// TIA Portal project "PROYECTO PICK AND PLACE FUNCIONA" (V17)

(* hardware
DEVICE "S7-1200 station_1"  S7-1200 Station
   slot 0: "Rack_0"  S7-1200 Rack  Rack  V1.0
   slot 1: "PLC_1"  CPU 1214C AC/DC/Rly  6ES7 214-1BG40-0XB0  V4.5
DEVICE "Estación PC"  SIMATIC PC station
   slot 0: "Estación PC"  Rail  SIMATIC PC-Station  V1.0
      slot 125: "Stationmanager"  Station_Manager  V6.0.4
   slot 1: "IE general_1"  IE General  IE_CP  V8.2.0
      slot 1: "PROFINET interface"  IEGeneral.Interface.8.2.0
   slot 2: "HMI_RT_2"  WinCC RT Advanced  6AV2 104-0xxxx-xxxx  17.0.0.0
      slot 33792: "Interfaz del equipo"  Host interface
*)

// ===== PLC "PLC_1"  CPU 1214C AC/DC/Rly =====

VAR_GLOBAL   // PLC tag table "Tabla de variables estándar"
   "System_Byte" AT %MB1 : Byte;
   "FirstScan" AT %M1.0 : Bool;
   "DiagStatusUpdate" AT %M1.1 : Bool;
   "AlwaysTRUE" AT %M1.2 : Bool;
   "AlwaysFALSE" AT %M1.3 : Bool;
   "Tag_1" AT %M700.3 : Bool;
   "Tag_2" AT %M700.4 : Bool;
   "Tag_3" AT %M900.0 : Bool;
   "Tag_4" AT %M900.1 : Bool;
   "Tag_5" AT %M900.5 : Bool;
   "MARCA_VENTOSA_V3" AT %M3000.0 : Bool;
   "Tag_6" AT %M8765.0 : Bool;
   "MARCA VACIA" AT %M3214.0 : Bool;
   "MARCA_VACIAA" AT %M4500.0 : Bool;
   "Tag_7" AT %MW5000 : Word;
   "Tag_8" AT %MD5000 : DWord;
   "RESET_CTU" AT %M5000.0 : Bool;
   "Tag_9" AT %MD5010 : DInt;
   "Tag_10" AT %M763.3 : Bool;
   "Tag_11" AT %M668.2 : Bool;
   "Tag_12" AT %M668.3 : Bool;
   "Tag_13" AT %M996.0 : Bool;
   "Tag_14" AT %M1200.0 : Bool;
   "Tag_15" AT %M1200.2 : Bool;
   "POSICIÓN 1" AT %M543.0 : Bool;
   "POSICIÓN 2" AT %M543.1 : Bool;
   "POSICIÓN 3" AT %M543.2 : Bool;
   "POSICIÓN 4" AT %M543.3 : Bool;
   "POSICIÓN 5" AT %M543.4 : Bool;
   "POSICIÓN 6" AT %M543.5 : Bool;
   "POSICIÓN 7" AT %M543.6 : Bool;
   "POSICIÓN 8" AT %M543.7 : Bool;
   "POSICIÓN 9" AT %M544.0 : Bool;
   "POSICIÓN 10" AT %M544.1 : Bool;
   "Tag_16" AT %M545.3 : Bool;
   "VALOR_PROCESO_ENTRADA" AT %QW15 : Int;
   "VALOR_PROCESO_SALIDA" AT %QW20 : Int;
END_VAR

VAR_GLOBAL   // PLC tag table "ENTRADAS Y SALIDAS"
   "PULSADOR_S1" AT %I0.0 : Bool;
   "PULSADOR_S2" AT %I0.1 : Bool;
   "SELECTOR_S3" AT %I0.2 : Bool;
   "PULSADOR_S4" AT %I0.3 : Bool;
   "DETECTOR_B1" AT %I0.4 : Bool;
   "DETECTOR_B2" AT %I0.5 : Bool;
   "DETECTOR_B3" AT %I0.6 : Bool;
   "DETECTOR_B4" AT %I0.7 : Bool;
   "DETECTOR_B5" AT %I1.0 : Bool;
   "E.VALVULA_MB1(B+)" AT %Q0.0 : Bool;
   "E.VALVULA_MB2(A+)" AT %Q0.1 : Bool;
   "CINTA1_KM1" AT %Q0.2 : Bool;
   "CINTA2_KM2" AT %Q0.3 : Bool;
   "VENTOSA_V1" AT %Q0.4 : Bool;
   "PILOTO_H2" AT %Q0.5 : Bool;
   "PILOTO_H1" AT %Q0.6 : Bool;
   "PILOTO_H3(AUTO)" AT %Q0.7 : Bool;
   "SELECTOR_S7" AT %I1.2 : Bool;
   "CINTA3_KM3" AT %Q1.0 : Bool;
   "CINTA4_KM4" AT %Q1.1 : Bool;
   "CINTA5_KM5" AT %Q1.2 : Bool;
   "CINTA6_KM6" AT %Q1.3 : Bool;
   "BARRERA1_KM7" AT %Q1.4 : Bool;
   "DETECTOR_B8=B3" AT %I1.4 : Bool;
   "DETECTOR C+_B9=B7" AT %I1.5 : Bool;
   "DETECTOR D+_B10=B6" AT %I1.6 : Bool;
   "DETECTOR_B11=B1" AT %I1.7 : Bool;
   "DETECTOR_B12=B4" AT %I2.0 : Bool;
   "DETECTOR_B13=B2" AT %I2.1 : Bool;
   "DETECTOR_B14=B5" AT %I2.2 : Bool;
   "BARRERA2_KM8" AT %Q1.5 : Bool;
   "PILOTO_H6(ROJO)" AT %Q2.0 : Bool;
   "PILOTO_H4(VERDE)" AT %Q2.1 : Bool;
   "PILOTO_H5(AMARILLO)" AT %Q2.2 : Bool;
   "M.MANUA2_S9" AT %I2.3 : Bool;
   "AUTO2_S10" AT %I2.4 : Bool;
   "MARCHA2_S5" AT %I2.5 : Bool;
   "PULSADOR_MANUAL_S6" AT %I2.6 : Bool;
   "PARO2_S8" AT %I2.7 : Bool;
   "PILOTO_H12=H1" AT %Q2.3 : Bool;
   "PILOTO_H7=H2" AT %Q2.4 : Bool;
   "PILOTO_H8=H3" AT %Q2.5 : Bool;
   "CINTA7_KM9=KM3" AT %Q2.6 : Bool;
   "PILOTO_H9=H4" AT %Q2.7 : Bool;
   "PILOTO_H10=H5" AT %Q3.0 : Bool;
   "PILOTO_H11=H6" AT %Q3.1 : Bool;
   "CILINDRO_C=A" AT %Q1.6 : Bool;
   "CILINDRO_D=B" AT %Q1.7 : Bool;
   "VENTOSA_V2" AT %Q3.2 : Bool;
   "FC1_E+" AT %I3.0 : Bool;
   "CILINDRO E" AT %Q5.0 : Bool;
   "FC2_E-" AT %I3.1 : Bool;
   "CÁMARA1_B15(AZUL)" AT %I3.2 : Bool;
   "CÁMARA2_B16(VERDE)" AT %I3.3 : Bool;
   "FC4_F+" AT %I3.4 : Bool;
   "FC5_G-" AT %I3.5 : Bool;
   "FC6_G+" AT %I3.6 : Bool;
   "FC3_F-" AT %I3.7 : Bool;
   "CILINDRO F" AT %Q5.1 : Bool;
   "CILINDRO G" AT %QD38 : DWord;
   "CINTA8_KM10" AT %Q3.3 : Bool;
   "PILOTOEMERGENCIA_H13" AT %Q3.4 : Bool;
   "SETAEMERGENCIA_S12" AT %I4.0 : Bool;
   "RESET1_S11" AT %I4.1 : Bool;
   "RESET2_S14" AT %I4.2 : Bool;
   "SETAEMERGENCIA2_S13" AT %I4.3 : Bool;
   "PILOTOEMERGENCIA2_H14" AT %Q3.5 : Bool;
   "DETECTOR_B15" AT %I4.4 : Bool;
   "ROBOT_OCUPADO_B16" AT %I4.5 : Bool;
   "ROBOT_ERROR_B17" AT %I4.6 : Bool;
   "ACTIVACIÓN_ROBOT" AT %Q3.6 : Bool;
   "DETECTOR_B21(INICIO P.AZUL)" AT %I4.7 : Bool;
   "DETECTOR_B22(FINAL P.AZUL)" AT %I5.0 : Bool;
   "CINTA9_KM11(BASE AZUL)" AT %Q3.7 : Bool;
   "CINTA10_KM12(BASE AZUL)" AT %Q4.0 : Bool;
   "CINTA11_KM13(BASE AZUL)" AT %Q4.1 : Bool;
   "BARRERA3_KM14(BASE AZUL)" AT %Q4.2 : Bool;
   "EJE_X1" AT %QD42 : Real;
   "EJE_Y1" AT %QD46 : Real;
   "EJE_Z1" AT %QD50 : Real;
   "VENTOSA_V3" AT %Q4.3 : Bool;
   "CINTA12_KM15(BASE VERDE)" AT %Q4.4 : Bool;
   "CINTA13_KM16(BASE VERDE)" AT %Q4.5 : Bool;
   "CINTA14_KM17(BASE VERDE)" AT %Q4.6 : Bool;
   "BARRERA4_KM18" AT %Q4.7 : Bool;
   "DETECTOR_B23(INICIO BASE VERDE)" AT %I5.1 : Bool;
   "DETECTOR_B24(FINAL BASE VERDE)" AT %I5.2 : Bool;
   "EJE_X2" AT %QD34 : Real;
   "EJE_Y2" AT %QD54 : Real;
   "EJE_Z2" AT %QD58 : Real;
   "VENTOSA_V4" AT %Q5.2 : Bool;
   "CINTA15_KM19" AT %Q5.3 : Bool;
   "CINTA16_KM20" AT %Q5.4 : Bool;
   "CINTA17_KM21" AT %Q5.5 : Bool;
   "CINTA18_KM22" AT %Q5.6 : Bool;
   "CINTA19_KM23" AT %Q5.7 : Bool;
   "CINTA20_KM24" AT %Q6.0 : Bool;
   "UÑASATRAS_KM25" AT %Q6.1 : Bool;
   "VAGÓN_ARRIBA_KM26" AT %Q6.2 : Bool;
   "SELECCION POSICIÓN" AT %QD30 : DInt;
   "DETECTOR_B25" AT %I5.3 : Bool;
   "DETECTOR_B26" AT %I5.4 : Bool;
   "SALIDA BASES" AT %Q6.3 : Bool;
   "SALIDA PALET_AZUL" AT %Q6.4 : Bool;
   "UÑAS_ALANTE_KM27" AT %Q6.5 : Bool;
   "CINTA21_KM28" AT %Q6.6 : Bool;
   "CINTA22_KM29" AT %Q6.7 : Bool;
   "CINTA23_KM30" AT %Q7.0 : Bool;
   "CINTA24_KM31" AT %Q7.1 : Bool;
   "CINTA25_KM32" AT %Q7.2 : Bool;
   "CINTA26_KM33" AT %Q7.3 : Bool;
   "DETECTOR_B27" AT %I5.5 : Bool;
   "DETECTOR_B28" AT %I5.6 : Bool;
   "SALIDA_PALET_VERDE" AT %Q7.4 : Bool;
   "VALOR_CONTADOR" AT %IW6 : Int;
   "MARCAA_VACIIA" AT %M730.0 : Bool;
END_VAR

VAR_GLOBAL   // PLC tag table "ETAPAS"
   "ETAPA_1" AT %M10.1 : Bool;
   "ETAPA_2" AT %M10.2 : Bool;
   "ETAPA_3" AT %M10.3 : Bool;
   "ETAPA_4" AT %M10.4 : Bool;
   "ETAPA_5" AT %M10.5 : Bool;
   "ETAPA_6" AT %M10.6 : Bool;
   "ETAPA_7" AT %M10.7 : Bool;
   "ETAPA_12" AT %M11.0 : Bool;
   "ETAPA_13" AT %M11.1 : Bool;
   "ETAPA_14" AT %M11.2 : Bool;
   "ETAPA_15" AT %M11.3 : Bool;
   "ETAPA_16" AT %M11.4 : Bool;
   "ETAPA_17" AT %M11.5 : Bool;
   "ETAPA_0" AT %M10.0 : Bool;
   "ETAPA_100" AT %M11.6 : Bool;
   "ETAPA_101" AT %M11.7 : Bool;
   "ETAPA_50" AT %M12.0 : Bool;
   "ETAPA_51" AT %M12.1 : Bool;
   "ETAPA_54" AT %M12.2 : Bool;
   "ETAPA_55" AT %M12.3 : Bool;
   "ETAPA_56" AT %M12.4 : Bool;
   "ETAPA_57" AT %M12.5 : Bool;
   "ETAPA_58" AT %M12.6 : Bool;
   "ETAPA_59" AT %M12.7 : Bool;
   "ETAPA_62" AT %M13.0 : Bool;
   "ETAPA_63" AT %M13.1 : Bool;
   "ETAPA_64" AT %M13.2 : Bool;
   "ETAPA_65" AT %M13.3 : Bool;
   "ETAPA_66" AT %M13.4 : Bool;
   "ETAPA_67" AT %M13.5 : Bool;
   "ETAPA_52" AT %M14.0 : Bool;
   "ETAPA_53" AT %M14.1 : Bool;
   "ETAPA_60" AT %M14.2 : Bool;
   "ETAPA_61" AT %M14.3 : Bool;
   "ETAPA_8" AT %M14.4 : Bool;
   "ETAPA_9" AT %M14.5 : Bool;
   "ETAPA_18" AT %M14.6 : Bool;
   "ETAPA_19" AT %M14.7 : Bool;
   "ETAPA_20" AT %M15.1 : Bool;
   "ETAPA_21" AT %M15.2 : Bool;
   "ETAPA _10" AT %M15.3 : Bool;
   "ETAPA_11" AT %M15.4 : Bool;
   "ETAPA_120" AT %M15.5 : Bool;
   "ETAPA_121" AT %M23.0 : Bool;
   "ETAPA_140" AT %M15.7 : Bool;
   "ETAPA_141" AT %M16.0 : Bool;
   "ETAPA_160" AT %M16.1 : Bool;
   "ETAPA_161" AT %M16.2 : Bool;
   "ETAPA_200" AT %M16.3 : Bool;
   "ETAPA_201" AT %M16.4 : Bool;
   "ETAPA_202" AT %M16.5 : Bool;
   "ETAPA_203" AT %M16.6 : Bool;
   "ETAPA_204" AT %M16.7 : Bool;
   "ETAPA_205" AT %M17.0 : Bool;
   "ETAPA_206" AT %M17.1 : Bool;
   "ETAPA_207" AT %M17.2 : Bool;
   "ETAPA_208" AT %M17.3 : Bool;
   "ETAPA_209" AT %M17.4 : Bool;
   "ETAPA_210" AT %M17.5 : Bool;
   "ETAPA_211" AT %M17.6 : Bool;
   "ETAPA_212" AT %M17.7 : Bool;
   "ETAPA_213" AT %M18.0 : Bool;
   "ETAPA_214" AT %M18.1 : Bool;
   "ETAPA_215" AT %M18.2 : Bool;
   "ETAPA_216" AT %M18.3 : Bool;
   "ETAPA_217" AT %M18.4 : Bool;
   "ETAPA_218" AT %M18.5 : Bool;
   "ETAPA_250" AT %M18.6 : Bool;
   "ETAPA_251" AT %M18.7 : Bool;
   "ETAPA_252" AT %M19.0 : Bool;
   "ETAPA_253" AT %M19.1 : Bool;
   "ETAPA_254" AT %M19.2 : Bool;
   "ETAPA_255" AT %M19.3 : Bool;
   "ETAPA_256" AT %M19.4 : Bool;
   "ETAPA_257" AT %M19.5 : Bool;
   "ETAPA_258" AT %M19.6 : Bool;
   "ETAPA_259" AT %M19.7 : Bool;
   "ETAPA_260" AT %M20.0 : Bool;
   "ETAPA_261" AT %M20.1 : Bool;
   "ETAPA_262" AT %M20.2 : Bool;
   "ETAPA_263" AT %M20.3 : Bool;
   "ETAPA_264" AT %M20.4 : Bool;
   "ETAPA_265" AT %M20.5 : Bool;
   "ETAPA_266" AT %M20.6 : Bool;
END_VAR

// folder: System blocks/Program resources

DATA_BLOCK "TEMPORIZADOR 1"   // DB1
{ S7_Optimized_Access := 'TRUE' }
AUTHOR : Simatic
FAMILY : IEC
NAME : IEC_TMR
VERSION : 1.0
// stored: InstanceOfName IEC_TIMER
"IEC_TIMER"
BEGIN
END_DATA_BLOCK

DATA_BLOCK "TEMPORIZADOR 2"   // DB2
{ S7_Optimized_Access := 'TRUE' }
AUTHOR : Simatic
FAMILY : IEC
NAME : IEC_TMR
VERSION : 1.0
// stored: InstanceOfName IEC_TIMER
"IEC_TIMER"
BEGIN
END_DATA_BLOCK

DATA_BLOCK "TEMPORIZADOR 3"   // DB3
{ S7_Optimized_Access := 'TRUE' }
AUTHOR : Simatic
FAMILY : IEC
NAME : IEC_TMR
VERSION : 1.0
// stored: InstanceOfName IEC_TIMER
"IEC_TIMER"
BEGIN
END_DATA_BLOCK

DATA_BLOCK "TEMPORIZADOR 4"   // DB4
{ S7_Optimized_Access := 'TRUE' }
AUTHOR : Simatic
FAMILY : IEC
NAME : IEC_TMR
VERSION : 1.0
// stored: InstanceOfName IEC_TIMER
"IEC_TIMER"
BEGIN
END_DATA_BLOCK

DATA_BLOCK "TEMPORIZADOR 5"   // DB5
{ S7_Optimized_Access := 'TRUE' }
AUTHOR : Simatic
FAMILY : IEC
NAME : IEC_TMR
VERSION : 1.0
// stored: InstanceOfName IEC_TIMER
"IEC_TIMER"
BEGIN
END_DATA_BLOCK

DATA_BLOCK "TEMPORIZADOR 6"   // DB6
{ S7_Optimized_Access := 'TRUE' }
AUTHOR : Simatic
FAMILY : IEC
NAME : IEC_TMR
VERSION : 1.0
// stored: InstanceOfName IEC_TIMER
"IEC_TIMER"
BEGIN
END_DATA_BLOCK

DATA_BLOCK "TEMPORIZADOR 10"   // DB7
{ S7_Optimized_Access := 'TRUE' }
AUTHOR : Simatic
FAMILY : IEC
NAME : IEC_TMR
VERSION : 1.0
// stored: InstanceOfName IEC_TIMER
"IEC_TIMER"
BEGIN
END_DATA_BLOCK

DATA_BLOCK "TEMPORIZADOR 8"   // DB8
{ S7_Optimized_Access := 'TRUE' }
AUTHOR : Simatic
FAMILY : IEC
NAME : IEC_TMR
VERSION : 1.0
// stored: InstanceOfName IEC_TIMER
"IEC_TIMER"
BEGIN
END_DATA_BLOCK

DATA_BLOCK "TEMPORIZADOR 13"   // DB9
{ S7_Optimized_Access := 'TRUE' }
AUTHOR : Simatic
FAMILY : IEC
NAME : IEC_TMR
VERSION : 1.0
// stored: InstanceOfName IEC_TIMER
"IEC_TIMER"
BEGIN
END_DATA_BLOCK

DATA_BLOCK "TEMPORIZADOR 15"   // DB10
{ S7_Optimized_Access := 'TRUE' }
AUTHOR : Simatic
FAMILY : IEC
NAME : IEC_TMR
VERSION : 1.0
// stored: InstanceOfName IEC_TIMER
"IEC_TIMER"
BEGIN
END_DATA_BLOCK

DATA_BLOCK "TEMPORIZADOR 11"   // DB11
{ S7_Optimized_Access := 'TRUE' }
AUTHOR : Simatic
FAMILY : IEC
NAME : IEC_TMR
VERSION : 1.0
// stored: InstanceOfName IEC_TIMER
"IEC_TIMER"
BEGIN
END_DATA_BLOCK

DATA_BLOCK "TEMPORIZADOR 14"   // DB12
{ S7_Optimized_Access := 'TRUE' }
AUTHOR : Simatic
FAMILY : IEC
NAME : IEC_TMR
VERSION : 1.0
// stored: InstanceOfName IEC_TIMER
"IEC_TIMER"
BEGIN
END_DATA_BLOCK

DATA_BLOCK "TEMPORIZADOR 7"   // DB13
{ S7_Optimized_Access := 'TRUE' }
AUTHOR : Simatic
FAMILY : IEC
NAME : IEC_TMR
VERSION : 1.0
// stored: InstanceOfName IEC_TIMER
"IEC_TIMER"
BEGIN
END_DATA_BLOCK

DATA_BLOCK "TEMPORIZADOR 16"   // DB14
{ S7_Optimized_Access := 'TRUE' }
AUTHOR : Simatic
FAMILY : IEC
NAME : IEC_TMR
VERSION : 1.0
// stored: InstanceOfName IEC_TIMER
"IEC_TIMER"
BEGIN
END_DATA_BLOCK

DATA_BLOCK "TEMPORIZADOR 17"   // DB15
{ S7_Optimized_Access := 'TRUE' }
AUTHOR : Simatic
FAMILY : IEC
NAME : IEC_TMR
VERSION : 1.0
// stored: InstanceOfName IEC_TIMER
"IEC_TIMER"
BEGIN
END_DATA_BLOCK

DATA_BLOCK "TEMPORIZADOR 18"   // DB16
{ S7_Optimized_Access := 'TRUE' }
AUTHOR : Simatic
FAMILY : IEC
NAME : IEC_TMR
VERSION : 1.0
// stored: InstanceOfName IEC_TIMER
"IEC_TIMER"
BEGIN
END_DATA_BLOCK

DATA_BLOCK "TEMPORIZADOR 19"   // DB17
{ S7_Optimized_Access := 'TRUE' }
AUTHOR : Simatic
FAMILY : IEC
NAME : IEC_TMR
VERSION : 1.0
// stored: InstanceOfName IEC_TIMER
"IEC_TIMER"
BEGIN
END_DATA_BLOCK

DATA_BLOCK "TEMPORIZADOR 20"   // DB18
{ S7_Optimized_Access := 'TRUE' }
AUTHOR : Simatic
FAMILY : IEC
NAME : IEC_TMR
VERSION : 1.0
// stored: InstanceOfName IEC_TIMER
"IEC_TIMER"
BEGIN
END_DATA_BLOCK

DATA_BLOCK "TEMPORIZADOR 21"   // DB19
{ S7_Optimized_Access := 'TRUE' }
AUTHOR : Simatic
FAMILY : IEC
NAME : IEC_TMR
VERSION : 1.0
// stored: InstanceOfName IEC_TIMER
"IEC_TIMER"
BEGIN
END_DATA_BLOCK

DATA_BLOCK "TEMPORIZADOR 22"   // DB20
{ S7_Optimized_Access := 'TRUE' }
AUTHOR : Simatic
FAMILY : IEC
NAME : IEC_TMR
VERSION : 1.0
// stored: InstanceOfName IEC_TIMER
"IEC_TIMER"
BEGIN
END_DATA_BLOCK

DATA_BLOCK "IEC_Timer_0_DB"   // DB21
{ S7_Optimized_Access := 'TRUE' }
AUTHOR : Simatic
FAMILY : IEC
NAME : IEC_TMR
VERSION : 1.0
// stored: InstanceOfName IEC_TIMER
"IEC_TIMER"
BEGIN
END_DATA_BLOCK

DATA_BLOCK "TEMPORIZADOR 23"   // DB22
{ S7_Optimized_Access := 'TRUE' }
AUTHOR : Simatic
FAMILY : IEC
NAME : IEC_TMR
VERSION : 1.0
// stored: InstanceOfName IEC_TIMER
"IEC_TIMER"
BEGIN
END_DATA_BLOCK

DATA_BLOCK "TEMPORIZADOR 24"   // DB23
{ S7_Optimized_Access := 'TRUE' }
AUTHOR : Simatic
FAMILY : IEC
NAME : IEC_TMR
VERSION : 1.0
// stored: InstanceOfName IEC_TIMER
"IEC_TIMER"
BEGIN
END_DATA_BLOCK

DATA_BLOCK "TEMPORIZADOR 25"   // DB24
{ S7_Optimized_Access := 'TRUE' }
AUTHOR : Simatic
FAMILY : IEC
NAME : IEC_TMR
VERSION : 1.0
// stored: InstanceOfName IEC_TIMER
"IEC_TIMER"
BEGIN
END_DATA_BLOCK

DATA_BLOCK "TEMPORIZADOR 26"   // DB25
{ S7_Optimized_Access := 'TRUE' }
AUTHOR : Simatic
FAMILY : IEC
NAME : IEC_TMR
VERSION : 1.0
// stored: InstanceOfName IEC_TIMER
"IEC_TIMER"
BEGIN
END_DATA_BLOCK

DATA_BLOCK "TEMPORIZADOR 27"   // DB26
{ S7_Optimized_Access := 'TRUE' }
AUTHOR : Simatic
FAMILY : IEC
NAME : IEC_TMR
VERSION : 1.0
// stored: InstanceOfName IEC_TIMER
"IEC_TIMER"
BEGIN
END_DATA_BLOCK

DATA_BLOCK "TEMPORIZADOR 28"   // DB27
{ S7_Optimized_Access := 'TRUE' }
AUTHOR : Simatic
FAMILY : IEC
NAME : IEC_TMR
VERSION : 1.0
// stored: InstanceOfName IEC_TIMER
"IEC_TIMER"
BEGIN
END_DATA_BLOCK

DATA_BLOCK "TEMPORIZADOR 29"   // DB28
{ S7_Optimized_Access := 'TRUE' }
AUTHOR : Simatic
FAMILY : IEC
NAME : IEC_TMR
VERSION : 1.0
// stored: InstanceOfName IEC_TIMER
"IEC_TIMER"
BEGIN
END_DATA_BLOCK

DATA_BLOCK "TEMPORIZADOR 30"   // DB29
{ S7_Optimized_Access := 'TRUE' }
AUTHOR : Simatic
FAMILY : IEC
NAME : IEC_TMR
VERSION : 1.0
// stored: InstanceOfName IEC_TIMER
"IEC_TIMER"
BEGIN
END_DATA_BLOCK

DATA_BLOCK "TEMPORIZADOR 31"   // DB30
{ S7_Optimized_Access := 'TRUE' }
AUTHOR : Simatic
FAMILY : IEC
NAME : IEC_TMR
VERSION : 1.0
// stored: InstanceOfName IEC_TIMER
"IEC_TIMER"
BEGIN
END_DATA_BLOCK

DATA_BLOCK "TEMPORIZADOR 32"   // DB31
{ S7_Optimized_Access := 'TRUE' }
AUTHOR : Simatic
FAMILY : IEC
NAME : IEC_TMR
VERSION : 1.0
// stored: InstanceOfName IEC_TIMER
"IEC_TIMER"
BEGIN
END_DATA_BLOCK

DATA_BLOCK "TEMPORIZADOR 33"   // DB32
{ S7_Optimized_Access := 'TRUE' }
AUTHOR : Simatic
FAMILY : IEC
NAME : IEC_TMR
VERSION : 1.0
// stored: InstanceOfName IEC_TIMER
"IEC_TIMER"
BEGIN
END_DATA_BLOCK

DATA_BLOCK "TEMPORIZADOR 34"   // DB33
{ S7_Optimized_Access := 'TRUE' }
AUTHOR : Simatic
FAMILY : IEC
NAME : IEC_TMR
VERSION : 1.0
// stored: InstanceOfName IEC_TIMER
"IEC_TIMER"
BEGIN
END_DATA_BLOCK

DATA_BLOCK "TEMPORIZADOR 35"   // DB34
{ S7_Optimized_Access := 'TRUE' }
AUTHOR : Simatic
FAMILY : IEC
NAME : IEC_TMR
VERSION : 1.0
// stored: InstanceOfName IEC_TIMER
"IEC_TIMER"
BEGIN
END_DATA_BLOCK

DATA_BLOCK "TEMPORIZADOR 36"   // DB35
{ S7_Optimized_Access := 'TRUE' }
AUTHOR : Simatic
FAMILY : IEC
NAME : IEC_TMR
VERSION : 1.0
// stored: InstanceOfName IEC_TIMER
"IEC_TIMER"
BEGIN
END_DATA_BLOCK

DATA_BLOCK "TEMPORIZADOR 37"   // DB36
{ S7_Optimized_Access := 'TRUE' }
AUTHOR : Simatic
FAMILY : IEC
NAME : IEC_TMR
VERSION : 1.0
// stored: InstanceOfName IEC_TIMER
"IEC_TIMER"
BEGIN
END_DATA_BLOCK

DATA_BLOCK "IEC_Timer_0_DB_1"   // DB37
{ S7_Optimized_Access := 'TRUE' }
AUTHOR : Simatic
FAMILY : IEC
NAME : IEC_TMR
VERSION : 1.0
// stored: InstanceOfName IEC_TIMER
"IEC_TIMER"
BEGIN
END_DATA_BLOCK

DATA_BLOCK "IEC_Counter_0_DB_1"   // DB38
{ S7_Optimized_Access := 'TRUE' }
AUTHOR : Simatic
FAMILY : IEC
NAME : CNTR
VERSION : 1.0
// stored: InstanceOfName IEC_COUNTER
"IEC_COUNTER"
BEGIN
END_DATA_BLOCK

DATA_BLOCK "IEC_Timer_0_DB_2"   // DB39
{ S7_Optimized_Access := 'TRUE' }
AUTHOR : Simatic
FAMILY : IEC
NAME : IEC_TMR
VERSION : 1.0
// stored: InstanceOfName IEC_TIMER
"IEC_TIMER"
BEGIN
END_DATA_BLOCK

DATA_BLOCK "IEC_Timer_0_DB_3"   // DB40
{ S7_Optimized_Access := 'TRUE' }
AUTHOR : Simatic
FAMILY : IEC
NAME : IEC_TMR
VERSION : 1.0
// stored: InstanceOfName IEC_TIMER
"IEC_TIMER"
BEGIN
END_DATA_BLOCK

DATA_BLOCK "TEMPORIZADOR 38"   // DB41
{ S7_Optimized_Access := 'TRUE' }
AUTHOR : Simatic
FAMILY : IEC
NAME : IEC_TMR
VERSION : 1.0
// stored: InstanceOfName IEC_TIMER
"IEC_TIMER"
BEGIN
END_DATA_BLOCK

DATA_BLOCK "TEMPORIZADOR 39"   // DB42
{ S7_Optimized_Access := 'TRUE' }
AUTHOR : Simatic
FAMILY : IEC
NAME : IEC_TMR
VERSION : 1.0
// stored: InstanceOfName IEC_TIMER
"IEC_TIMER"
BEGIN
END_DATA_BLOCK

DATA_BLOCK "IEC_Timer_0_DB_4"   // DB43
{ S7_Optimized_Access := 'TRUE' }
AUTHOR : Simatic
FAMILY : IEC
NAME : IEC_TMR
VERSION : 1.0
// stored: InstanceOfName IEC_TIMER
"IEC_TIMER"
BEGIN
END_DATA_BLOCK

DATA_BLOCK "IEC_Timer_0_DB_5"   // DB44
{ S7_Optimized_Access := 'TRUE' }
AUTHOR : Simatic
FAMILY : IEC
NAME : IEC_TMR
VERSION : 1.0
// stored: InstanceOfName IEC_TIMER
"IEC_TIMER"
BEGIN
END_DATA_BLOCK

DATA_BLOCK "TEMPORIZADOR 40"   // DB45
{ S7_Optimized_Access := 'TRUE' }
AUTHOR : Simatic
FAMILY : IEC
NAME : IEC_TMR
VERSION : 1.0
// stored: InstanceOfName IEC_TIMER
"IEC_TIMER"
BEGIN
END_DATA_BLOCK

DATA_BLOCK "TEMPORIZADOR 41"   // DB46
{ S7_Optimized_Access := 'TRUE' }
AUTHOR : Simatic
FAMILY : IEC
NAME : IEC_TMR
VERSION : 1.0
// stored: InstanceOfName IEC_TIMER
"IEC_TIMER"
BEGIN
END_DATA_BLOCK

DATA_BLOCK "TEMPORIZADOR 42"   // DB47
{ S7_Optimized_Access := 'TRUE' }
AUTHOR : Simatic
FAMILY : IEC
NAME : IEC_TMR
VERSION : 1.0
// stored: InstanceOfName IEC_TIMER
"IEC_TIMER"
BEGIN
END_DATA_BLOCK

DATA_BLOCK "TEMPORIZADOR 43"   // DB48
{ S7_Optimized_Access := 'TRUE' }
AUTHOR : Simatic
FAMILY : IEC
NAME : IEC_TMR
VERSION : 1.0
// stored: InstanceOfName IEC_TIMER
"IEC_TIMER"
BEGIN
END_DATA_BLOCK

DATA_BLOCK "TEMPORIZADOR 44"   // DB49
{ S7_Optimized_Access := 'TRUE' }
AUTHOR : Simatic
FAMILY : IEC
NAME : IEC_TMR
VERSION : 1.0
// stored: InstanceOfName IEC_TIMER
"IEC_TIMER"
BEGIN
END_DATA_BLOCK

DATA_BLOCK "TEMPORIZADOR 45"   // DB50
{ S7_Optimized_Access := 'TRUE' }
AUTHOR : Simatic
FAMILY : IEC
NAME : IEC_TMR
VERSION : 1.0
// stored: InstanceOfName IEC_TIMER
"IEC_TIMER"
BEGIN
END_DATA_BLOCK

// folder: (top level)

FUNCTION "FC_SECUENCIA SALIDA PARTE 1" : Void   // FC1, LAD
TITLE = PROGRAMACIÓN DEL PROCESO INDUSTRIAL
{ S7_Optimized_Access := 'TRUE' }
VERSION : 0.1
// ESTE BLOQUE MUESTRA LA PROGRAMACIÓN DE LA SECUENCIA DEL PROCESO INDUSTRIAL, DESDE QUE SALE DEL ROBOT HASTA QUE PASA LAS CÁMARAS DE VISIÓN DE COLORES
   VAR_TEMP   // added for the SCL form of the ladder/FBD networks
      _w1 : Bool;
      _w2 : Bool;
      _w3 : Bool;
      _w4 : Bool;
      _w5 : Bool;
   END_VAR
BEGIN

REGION Network 1: SET EN LA ETAPA 0
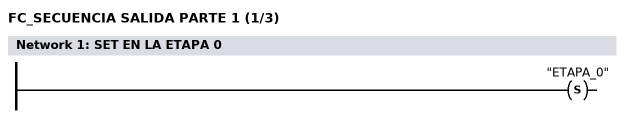
   RUNG wire#powerrail
      S_Coil( "ETAPA_0" )
   END_RUNG
   // the same network as SCL:
   "ETAPA_0" := TRUE;
END_REGION

REGION Network 2: PROGRAMACIÓN DE LA SECUENCIA EN MODO AUTOMÁTICO
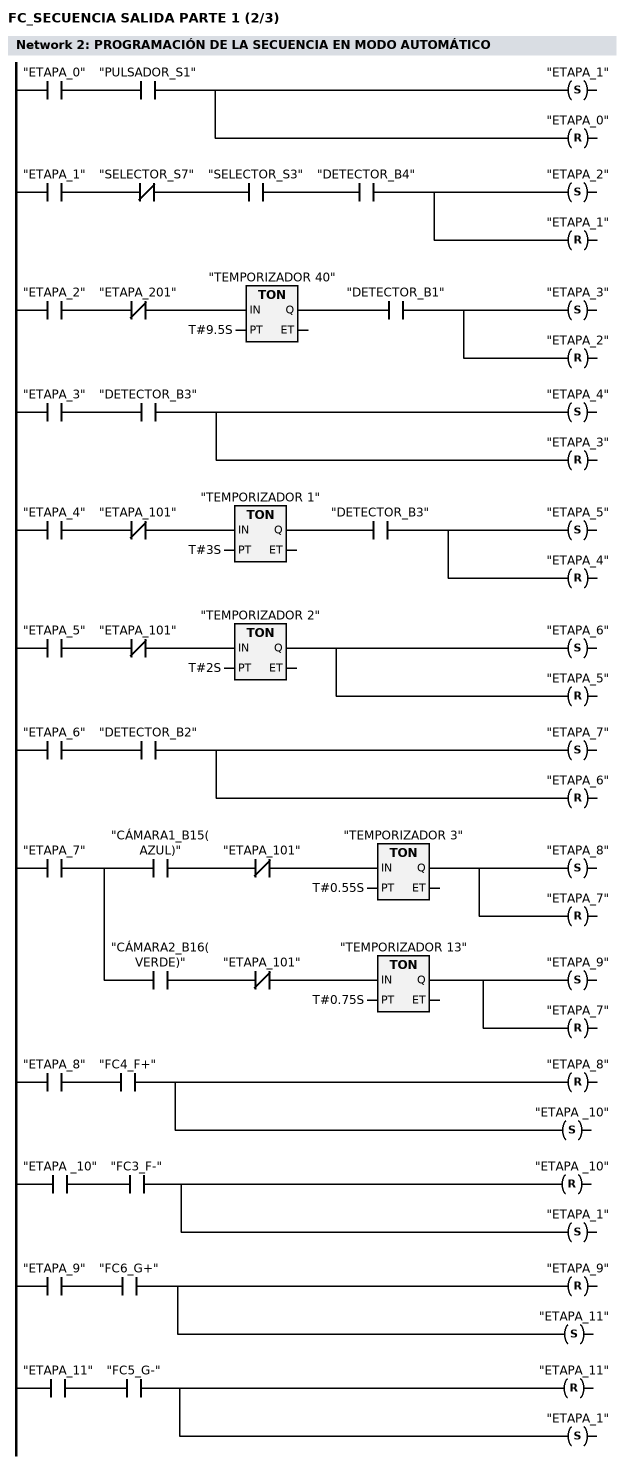
   IF "ETAPA_0" AND "PULSADOR_S1" THEN
       "ETAPA_1" := TRUE;
       "ETAPA_0" := FALSE;
   END_IF;
   IF "ETAPA_1" AND NOT "SELECTOR_S7" AND "SELECTOR_S3" AND "DETECTOR_B4" THEN
       "ETAPA_2" := TRUE;
       "ETAPA_1" := FALSE;
   END_IF;
   "TEMPORIZADOR 40".TON(IN := "ETAPA_2" AND NOT "ETAPA_201", PT := T#9.5S);
   IF "TEMPORIZADOR 40".Q AND "DETECTOR_B1" THEN
       "ETAPA_3" := TRUE;
       "ETAPA_2" := FALSE;
   END_IF;
   IF "ETAPA_3" AND "DETECTOR_B3" THEN
       "ETAPA_4" := TRUE;
       "ETAPA_3" := FALSE;
   END_IF;
   "TEMPORIZADOR 1".TON(IN := "ETAPA_4" AND NOT "ETAPA_101", PT := T#3S);
   IF "TEMPORIZADOR 1".Q AND "DETECTOR_B3" THEN
       "ETAPA_5" := TRUE;
       "ETAPA_4" := FALSE;
   END_IF;
   "TEMPORIZADOR 2".TON(IN := "ETAPA_5" AND NOT "ETAPA_101", PT := T#2S);
   IF "TEMPORIZADOR 2".Q THEN
       "ETAPA_6" := TRUE;
       "ETAPA_5" := FALSE;
   END_IF;
   IF "ETAPA_6" AND "DETECTOR_B2" THEN
       "ETAPA_7" := TRUE;
       "ETAPA_6" := FALSE;
   END_IF;
   "TEMPORIZADOR 3".TON(IN := "ETAPA_7" AND "CÁMARA1_B15(AZUL)" AND NOT "ETAPA_101", PT := T#0.55S);
   IF "TEMPORIZADOR 3".Q THEN "ETAPA_8" := TRUE; END_IF;
   #_w1 := "ETAPA_7";
   IF "TEMPORIZADOR 3".Q THEN "ETAPA_7" := FALSE; END_IF;
   "TEMPORIZADOR 13".TON(IN := #_w1 AND "CÁMARA2_B16(VERDE)" AND NOT "ETAPA_101", PT := T#0.75S);
   IF "TEMPORIZADOR 13".Q THEN
       "ETAPA_9" := TRUE;
       "ETAPA_7" := FALSE;
   END_IF;
   #_w2 := "ETAPA_8" AND "FC4_F+";
   IF #_w2 THEN
       "ETAPA_8" := FALSE;
       "ETAPA _10" := TRUE;
   END_IF;
   #_w3 := "ETAPA _10" AND "FC3_F-";
   IF #_w3 THEN
       "ETAPA _10" := FALSE;
       "ETAPA_1" := TRUE;
   END_IF;
   #_w4 := "ETAPA_9" AND "FC6_G+";
   IF #_w4 THEN
       "ETAPA_9" := FALSE;
       "ETAPA_11" := TRUE;
   END_IF;
   #_w5 := "ETAPA_11" AND "FC5_G-";
   IF #_w5 THEN
       "ETAPA_11" := FALSE;
       "ETAPA_1" := TRUE;
   END_IF;
END_REGION

REGION Network 3: PROGRAMACIÓN DE LA SECUENCIA EN MODO MANUAL
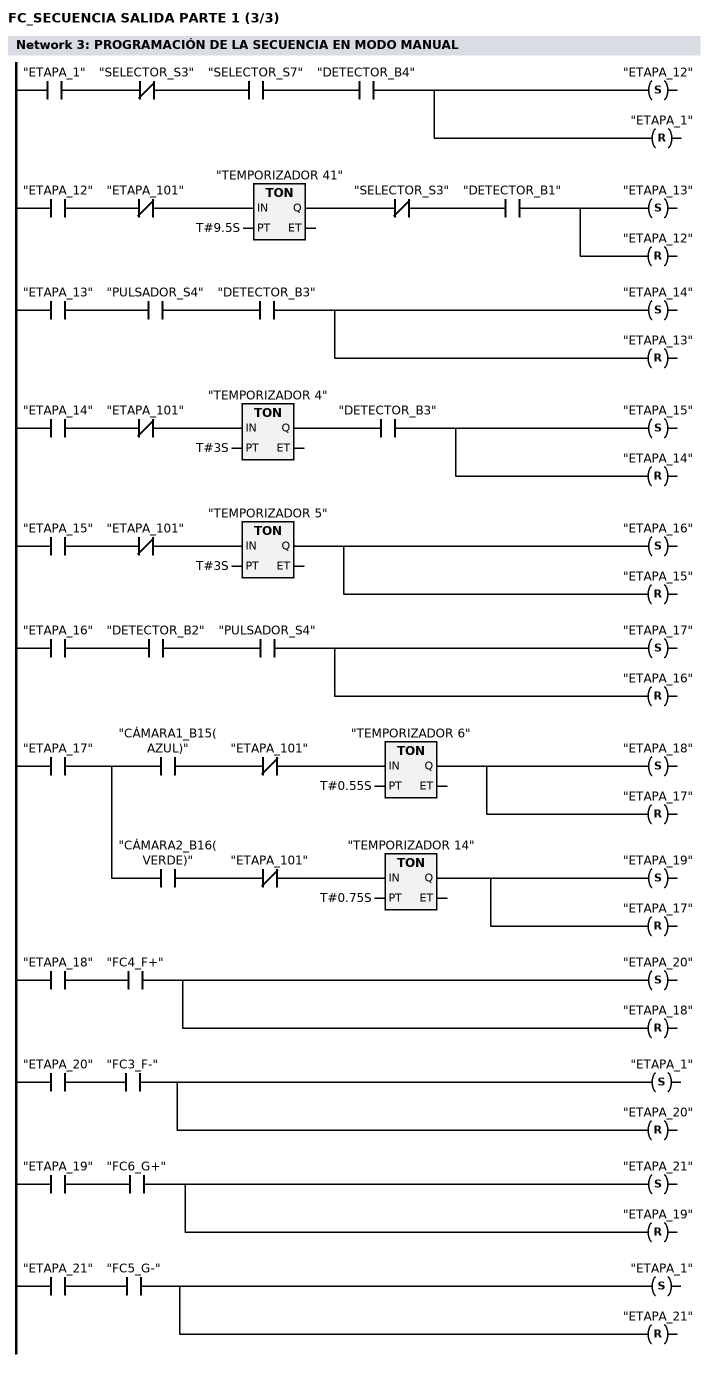
   IF "ETAPA_1" AND NOT "SELECTOR_S3" AND "SELECTOR_S7" AND "DETECTOR_B4" THEN
       "ETAPA_12" := TRUE;
       "ETAPA_1" := FALSE;
   END_IF;
   "TEMPORIZADOR 41".TON(IN := "ETAPA_12" AND NOT "ETAPA_101", PT := T#9.5S);
   IF "TEMPORIZADOR 41".Q AND NOT "SELECTOR_S3" AND "DETECTOR_B1" THEN
       "ETAPA_13" := TRUE;
       "ETAPA_12" := FALSE;
   END_IF;
   IF "ETAPA_13" AND "PULSADOR_S4" AND "DETECTOR_B3" THEN
       "ETAPA_14" := TRUE;
       "ETAPA_13" := FALSE;
   END_IF;
   "TEMPORIZADOR 4".TON(IN := "ETAPA_14" AND NOT "ETAPA_101", PT := T#3S);
   IF "TEMPORIZADOR 4".Q AND "DETECTOR_B3" THEN
       "ETAPA_15" := TRUE;
       "ETAPA_14" := FALSE;
   END_IF;
   "TEMPORIZADOR 5".TON(IN := "ETAPA_15" AND NOT "ETAPA_101", PT := T#3S);
   IF "TEMPORIZADOR 5".Q THEN
       "ETAPA_16" := TRUE;
       "ETAPA_15" := FALSE;
   END_IF;
   IF "ETAPA_16" AND "DETECTOR_B2" AND "PULSADOR_S4" THEN
       "ETAPA_17" := TRUE;
       "ETAPA_16" := FALSE;
   END_IF;
   "TEMPORIZADOR 6".TON(IN := "ETAPA_17" AND "CÁMARA1_B15(AZUL)" AND NOT "ETAPA_101", PT := T#0.55S);
   IF "TEMPORIZADOR 6".Q THEN "ETAPA_18" := TRUE; END_IF;
   #_w1 := "ETAPA_17";
   IF "TEMPORIZADOR 6".Q THEN "ETAPA_17" := FALSE; END_IF;
   "TEMPORIZADOR 14".TON(IN := #_w1 AND "CÁMARA2_B16(VERDE)" AND NOT "ETAPA_101", PT := T#0.75S);
   IF "TEMPORIZADOR 14".Q THEN
       "ETAPA_19" := TRUE;
       "ETAPA_17" := FALSE;
   END_IF;
   IF "ETAPA_18" AND "FC4_F+" THEN
       "ETAPA_20" := TRUE;
       "ETAPA_18" := FALSE;
   END_IF;
   IF "ETAPA_20" AND "FC3_F-" THEN
       "ETAPA_1" := TRUE;
       "ETAPA_20" := FALSE;
   END_IF;
   IF "ETAPA_19" AND "FC6_G+" THEN
       "ETAPA_21" := TRUE;
       "ETAPA_19" := FALSE;
   END_IF;
   IF "ETAPA_21" AND "FC5_G-" THEN
       "ETAPA_1" := TRUE;
       "ETAPA_21" := FALSE;
   END_IF;
END_REGION
END_FUNCTION

FUNCTION "FC_BOBINAS SALIDA PARTE 1" : Void   // FC2, LAD
TITLE = EN ESTE BLOQUE VEMOS LA ACCIÓN QUE HACE CADA ETAPA
{ S7_Optimized_Access := 'TRUE' }
VERSION : 0.1
// EN ESTE BLOQUE SE ENCUENTRA LA ASIGNACIÓN DE CADA ETAPA CON EL ACTUADOR QUE CORRESPONDE, DESDE LA SALIDA DEL ROBOT HASTA PASAR LAS CÁMARAS DE VISIÓN DE COLORES
BEGIN

REGION Network 1: ASIGNACIÓN DE LAS BOBINAS CON SU CORRESPONDIENTE ACTUADOR; PROCESO DE SALIDA
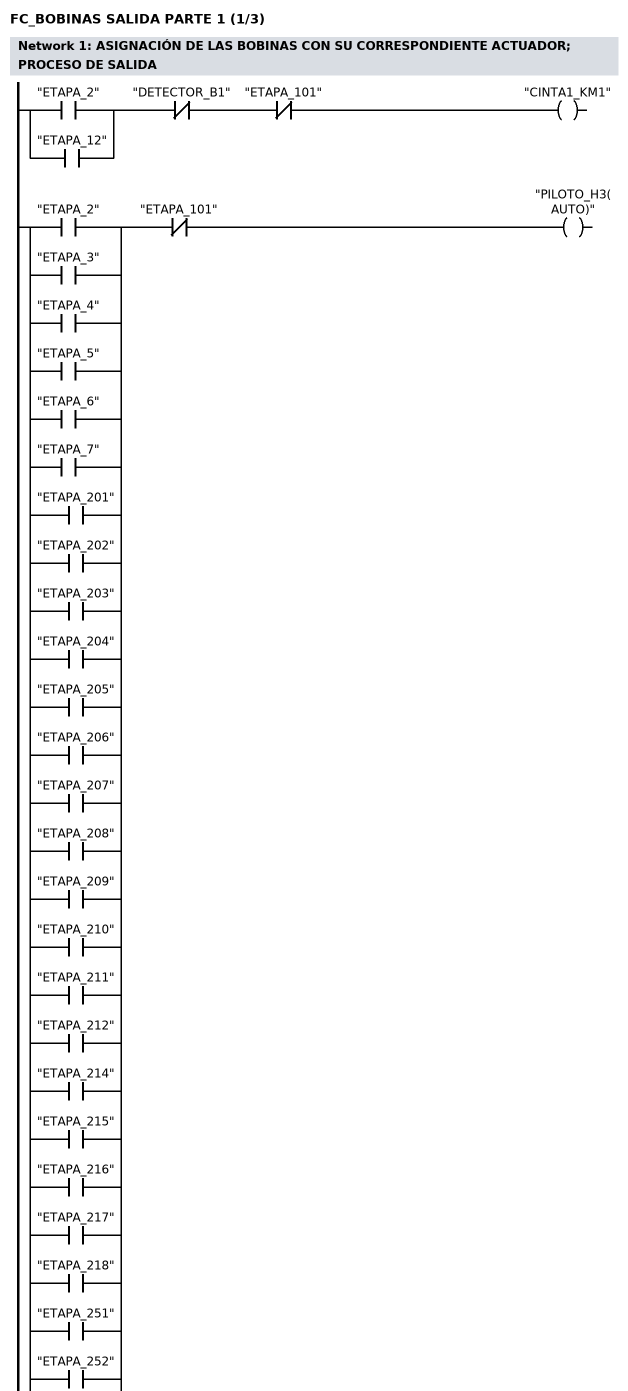
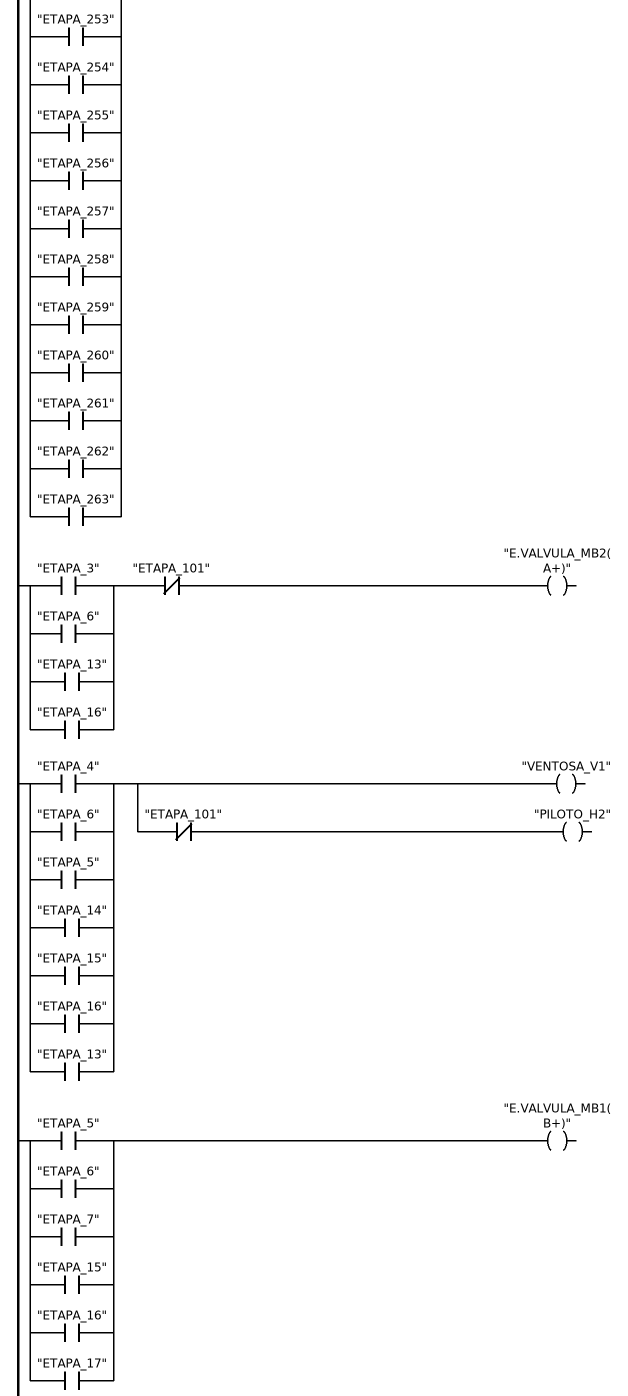
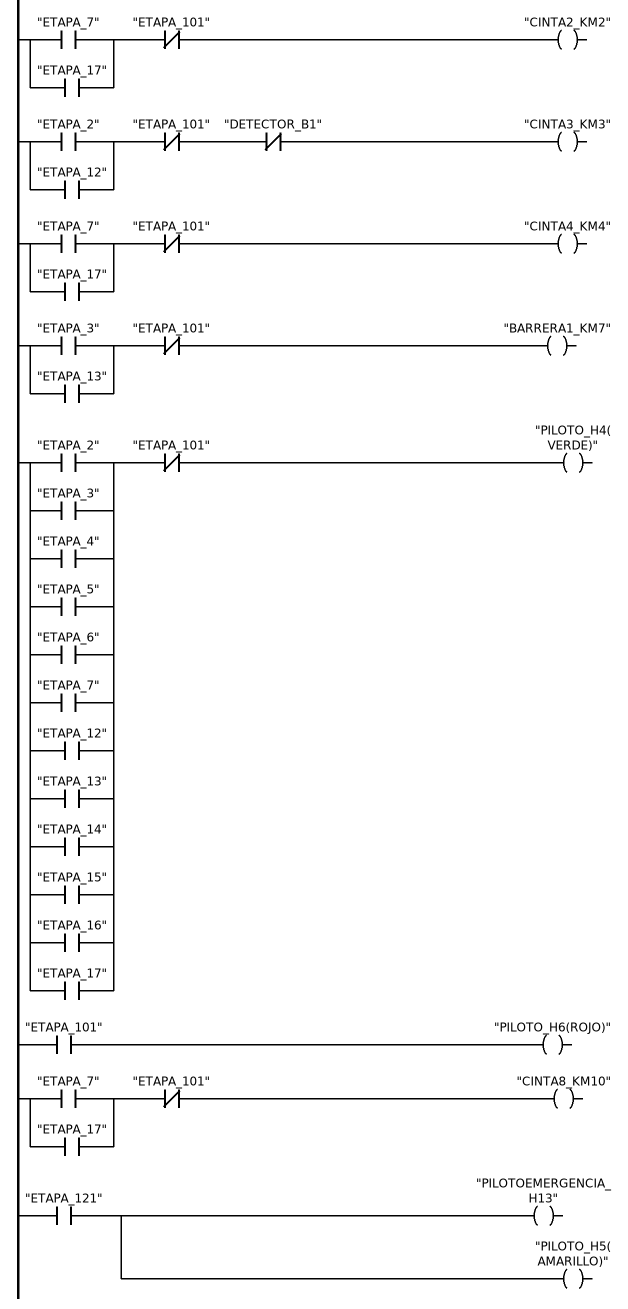
   RUNG wire#powerrail
      Contact( "ETAPA_2" )
      wire#w1
      I_Contact( "DETECTOR_B1" )
      I_Contact( "ETAPA_101" )
      Coil( "CINTA1_KM1" )
   END_RUNG
   RUNG wire#powerrail
      Contact( "ETAPA_12" )
   END_RUNG wire#w1
   RUNG wire#powerrail
      Contact( "ETAPA_2" )
      wire#w2
      I_Contact( "ETAPA_101" )
      Coil( "PILOTO_H3(AUTO)" )
   END_RUNG
   RUNG wire#powerrail
      Contact( "ETAPA_3" )
   END_RUNG wire#w2
   RUNG wire#powerrail
      Contact( "ETAPA_4" )
   END_RUNG wire#w2
   RUNG wire#powerrail
      Contact( "ETAPA_5" )
   END_RUNG wire#w2
   RUNG wire#powerrail
      Contact( "ETAPA_6" )
   END_RUNG wire#w2
   RUNG wire#powerrail
      Contact( "ETAPA_7" )
   END_RUNG wire#w2
   RUNG wire#powerrail
      Contact( "ETAPA_201" )
   END_RUNG wire#w2
   RUNG wire#powerrail
      Contact( "ETAPA_202" )
   END_RUNG wire#w2
   RUNG wire#powerrail
      Contact( "ETAPA_203" )
   END_RUNG wire#w2
   RUNG wire#powerrail
      Contact( "ETAPA_204" )
   END_RUNG wire#w2
   RUNG wire#powerrail
      Contact( "ETAPA_205" )
   END_RUNG wire#w2
   RUNG wire#powerrail
      Contact( "ETAPA_206" )
   END_RUNG wire#w2
   RUNG wire#powerrail
      Contact( "ETAPA_207" )
   END_RUNG wire#w2
   RUNG wire#powerrail
      Contact( "ETAPA_208" )
   END_RUNG wire#w2
   RUNG wire#powerrail
      Contact( "ETAPA_209" )
   END_RUNG wire#w2
   RUNG wire#powerrail
      Contact( "ETAPA_210" )
   END_RUNG wire#w2
   RUNG wire#powerrail
      Contact( "ETAPA_211" )
   END_RUNG wire#w2
   RUNG wire#powerrail
      Contact( "ETAPA_212" )
   END_RUNG wire#w2
   RUNG wire#powerrail
      Contact( "ETAPA_214" )
   END_RUNG wire#w2
   RUNG wire#powerrail
      Contact( "ETAPA_215" )
   END_RUNG wire#w2
   RUNG wire#powerrail
      Contact( "ETAPA_216" )
   END_RUNG wire#w2
   RUNG wire#powerrail
      Contact( "ETAPA_217" )
   END_RUNG wire#w2
   RUNG wire#powerrail
      Contact( "ETAPA_218" )
   END_RUNG wire#w2
   RUNG wire#powerrail
      Contact( "ETAPA_251" )
   END_RUNG wire#w2
   RUNG wire#powerrail
      Contact( "ETAPA_252" )
   END_RUNG wire#w2
   RUNG wire#powerrail
      Contact( "ETAPA_253" )
   END_RUNG wire#w2
   RUNG wire#powerrail
      Contact( "ETAPA_254" )
   END_RUNG wire#w2
   RUNG wire#powerrail
      Contact( "ETAPA_255" )
   END_RUNG wire#w2
   RUNG wire#powerrail
      Contact( "ETAPA_256" )
   END_RUNG wire#w2
   RUNG wire#powerrail
      Contact( "ETAPA_257" )
   END_RUNG wire#w2
   RUNG wire#powerrail
      Contact( "ETAPA_258" )
   END_RUNG wire#w2
   RUNG wire#powerrail
      Contact( "ETAPA_259" )
   END_RUNG wire#w2
   RUNG wire#powerrail
      Contact( "ETAPA_260" )
   END_RUNG wire#w2
   RUNG wire#powerrail
      Contact( "ETAPA_261" )
   END_RUNG wire#w2
   RUNG wire#powerrail
      Contact( "ETAPA_262" )
   END_RUNG wire#w2
   RUNG wire#powerrail
      Contact( "ETAPA_263" )
   END_RUNG wire#w2
   RUNG wire#powerrail
      Contact( "ETAPA_3" )
      wire#w3
      I_Contact( "ETAPA_101" )
      Coil( "E.VALVULA_MB2(A+)" )
   END_RUNG
   RUNG wire#powerrail
      Contact( "ETAPA_6" )
   END_RUNG wire#w3
   RUNG wire#powerrail
      Contact( "ETAPA_13" )
   END_RUNG wire#w3
   RUNG wire#powerrail
      Contact( "ETAPA_16" )
   END_RUNG wire#w3
   RUNG wire#powerrail
      Contact( "ETAPA_4" )
      wire#w4
      Coil( "VENTOSA_V1" )
   END_RUNG
   RUNG wire#powerrail
      Contact( "ETAPA_6" )
   END_RUNG wire#w4
   RUNG wire#powerrail
      Contact( "ETAPA_5" )
   END_RUNG wire#w4
   RUNG wire#powerrail
      Contact( "ETAPA_14" )
   END_RUNG wire#w4
   RUNG wire#powerrail
      Contact( "ETAPA_15" )
   END_RUNG wire#w4
   RUNG wire#powerrail
      Contact( "ETAPA_16" )
   END_RUNG wire#w4
   RUNG wire#powerrail
      Contact( "ETAPA_13" )
   END_RUNG wire#w4
   RUNG wire#w4
      I_Contact( "ETAPA_101" )
      Coil( "PILOTO_H2" )
   END_RUNG
   RUNG wire#powerrail
      Contact( "ETAPA_5" )
      wire#w5
      Coil( "E.VALVULA_MB1(B+)" )
   END_RUNG
   RUNG wire#powerrail
      Contact( "ETAPA_6" )
   END_RUNG wire#w5
   RUNG wire#powerrail
      Contact( "ETAPA_7" )
   END_RUNG wire#w5
   RUNG wire#powerrail
      Contact( "ETAPA_15" )
   END_RUNG wire#w5
   RUNG wire#powerrail
      Contact( "ETAPA_16" )
   END_RUNG wire#w5
   RUNG wire#powerrail
      Contact( "ETAPA_17" )
   END_RUNG wire#w5
   RUNG wire#powerrail
      Contact( "ETAPA_7" )
      wire#w6
      I_Contact( "ETAPA_101" )
      Coil( "CINTA2_KM2" )
   END_RUNG
   RUNG wire#powerrail
      Contact( "ETAPA_17" )
   END_RUNG wire#w6
   RUNG wire#powerrail
      Contact( "ETAPA_2" )
      wire#w7
      I_Contact( "ETAPA_101" )
      I_Contact( "DETECTOR_B1" )
      Coil( "CINTA3_KM3" )
   END_RUNG
   RUNG wire#powerrail
      Contact( "ETAPA_12" )
   END_RUNG wire#w7
   RUNG wire#powerrail
      Contact( "ETAPA_7" )
      wire#w8
      I_Contact( "ETAPA_101" )
      Coil( "CINTA4_KM4" )
   END_RUNG
   RUNG wire#powerrail
      Contact( "ETAPA_17" )
   END_RUNG wire#w8
   RUNG wire#powerrail
      Contact( "ETAPA_3" )
      wire#w9
      I_Contact( "ETAPA_101" )
      Coil( "BARRERA1_KM7" )
   END_RUNG
   RUNG wire#powerrail
      Contact( "ETAPA_13" )
   END_RUNG wire#w9
   RUNG wire#powerrail
      Contact( "ETAPA_2" )
      wire#w10
      I_Contact( "ETAPA_101" )
      Coil( "PILOTO_H4(VERDE)" )
   END_RUNG
   RUNG wire#powerrail
      Contact( "ETAPA_3" )
   END_RUNG wire#w10
   RUNG wire#powerrail
      Contact( "ETAPA_4" )
   END_RUNG wire#w10
   RUNG wire#powerrail
      Contact( "ETAPA_5" )
   END_RUNG wire#w10
   RUNG wire#powerrail
      Contact( "ETAPA_6" )
   END_RUNG wire#w10
   RUNG wire#powerrail
      Contact( "ETAPA_7" )
   END_RUNG wire#w10
   RUNG wire#powerrail
      Contact( "ETAPA_12" )
   END_RUNG wire#w10
   RUNG wire#powerrail
      Contact( "ETAPA_13" )
   END_RUNG wire#w10
   RUNG wire#powerrail
      Contact( "ETAPA_14" )
   END_RUNG wire#w10
   RUNG wire#powerrail
      Contact( "ETAPA_15" )
   END_RUNG wire#w10
   RUNG wire#powerrail
      Contact( "ETAPA_16" )
   END_RUNG wire#w10
   RUNG wire#powerrail
      Contact( "ETAPA_17" )
   END_RUNG wire#w10
   RUNG wire#powerrail
      Contact( "ETAPA_101" )
      Coil( "PILOTO_H6(ROJO)" )
   END_RUNG
   RUNG wire#powerrail
      Contact( "ETAPA_7" )
      wire#w11
      I_Contact( "ETAPA_101" )
      Coil( "CINTA8_KM10" )
   END_RUNG
   RUNG wire#powerrail
      Contact( "ETAPA_17" )
   END_RUNG wire#w11
   RUNG wire#powerrail
      Contact( "ETAPA_121" )
      wire#w12
      Coil( "PILOTOEMERGENCIA_H13" )
   END_RUNG
   RUNG wire#w12
      Coil( "PILOTO_H5(AMARILLO)" )
   END_RUNG
   // the same network as SCL:
   "CINTA1_KM1" := ("ETAPA_2" OR "ETAPA_12") AND NOT "DETECTOR_B1" AND NOT "ETAPA_101";
   "PILOTO_H3(AUTO)" := ("ETAPA_2" OR "ETAPA_3" OR "ETAPA_4" OR "ETAPA_5" OR "ETAPA_6" OR "ETAPA_7" OR "ETAPA_201" OR "ETAPA_202" OR "ETAPA_203" OR "ETAPA_204" OR "ETAPA_205" OR "ETAPA_206" OR "ETAPA_207" OR "ETAPA_208" OR "ETAPA_209" OR "ETAPA_210" OR "ETAPA_211" OR "ETAPA_212" OR "ETAPA_214" OR "ETAPA_215" OR "ETAPA_216" OR "ETAPA_217" OR "ETAPA_218" OR "ETAPA_251" OR "ETAPA_252" OR "ETAPA_253" OR "ETAPA_254" OR "ETAPA_255" OR "ETAPA_256" OR "ETAPA_257" OR "ETAPA_258" OR "ETAPA_259" OR "ETAPA_260" OR "ETAPA_261" OR "ETAPA_262" OR "ETAPA_263") AND NOT "ETAPA_101";
   "E.VALVULA_MB2(A+)" := ("ETAPA_3" OR "ETAPA_6" OR "ETAPA_13" OR "ETAPA_16") AND NOT "ETAPA_101";
   "VENTOSA_V1" := "ETAPA_4" OR "ETAPA_6" OR "ETAPA_5" OR "ETAPA_14" OR "ETAPA_15" OR "ETAPA_16" OR "ETAPA_13";
   "PILOTO_H2" := "VENTOSA_V1" AND NOT "ETAPA_101";
   "E.VALVULA_MB1(B+)" := "ETAPA_5" OR "ETAPA_6" OR "ETAPA_7" OR "ETAPA_15" OR "ETAPA_16" OR "ETAPA_17";
   "CINTA2_KM2" := ("ETAPA_7" OR "ETAPA_17") AND NOT "ETAPA_101";
   "CINTA3_KM3" := ("ETAPA_2" OR "ETAPA_12") AND NOT "ETAPA_101" AND NOT "DETECTOR_B1";
   "CINTA4_KM4" := ("ETAPA_7" OR "ETAPA_17") AND NOT "ETAPA_101";
   "BARRERA1_KM7" := ("ETAPA_3" OR "ETAPA_13") AND NOT "ETAPA_101";
   "PILOTO_H4(VERDE)" := ("ETAPA_2" OR "ETAPA_3" OR "ETAPA_4" OR "ETAPA_5" OR "ETAPA_6" OR "ETAPA_7" OR "ETAPA_12" OR "ETAPA_13" OR "ETAPA_14" OR "ETAPA_15" OR "ETAPA_16" OR "ETAPA_17") AND NOT "ETAPA_101";
   "PILOTO_H6(ROJO)" := "ETAPA_101";
   "CINTA8_KM10" := ("ETAPA_7" OR "ETAPA_17") AND NOT "ETAPA_101";
   "PILOTOEMERGENCIA_H13" := "ETAPA_121";
   "PILOTO_H5(AMARILLO)" := "ETAPA_121";
END_REGION

REGION Network 2
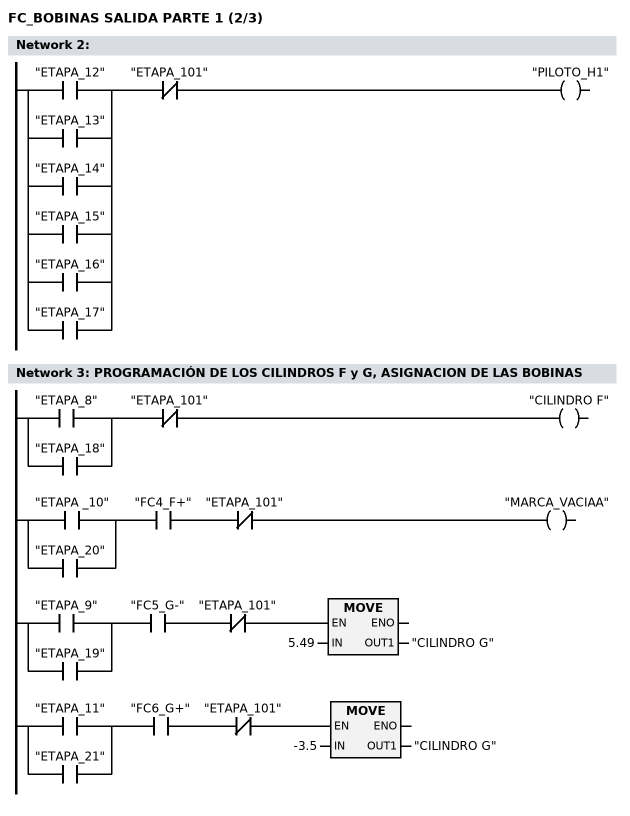
   RUNG wire#powerrail
      Contact( "ETAPA_12" )
      wire#w1
      I_Contact( "ETAPA_101" )
      Coil( "PILOTO_H1" )
   END_RUNG
   RUNG wire#powerrail
      Contact( "ETAPA_13" )
   END_RUNG wire#w1
   RUNG wire#powerrail
      Contact( "ETAPA_14" )
   END_RUNG wire#w1
   RUNG wire#powerrail
      Contact( "ETAPA_15" )
   END_RUNG wire#w1
   RUNG wire#powerrail
      Contact( "ETAPA_16" )
   END_RUNG wire#w1
   RUNG wire#powerrail
      Contact( "ETAPA_17" )
   END_RUNG wire#w1
   // the same network as SCL:
   "PILOTO_H1" := ("ETAPA_12" OR "ETAPA_13" OR "ETAPA_14" OR "ETAPA_15" OR "ETAPA_16" OR "ETAPA_17") AND NOT "ETAPA_101";
END_REGION

REGION Network 3: PROGRAMACIÓN DE LOS CILINDROS F y G, ASIGNACION DE LAS BOBINAS
   RUNG wire#powerrail
      Contact( "ETAPA_8" )
      wire#w1
      I_Contact( "ETAPA_101" )
      Coil( "CILINDRO F" )
   END_RUNG
   RUNG wire#powerrail
      Contact( "ETAPA_18" )
   END_RUNG wire#w1
   RUNG wire#powerrail
      Contact( "ETAPA _10" )
      wire#w2
      Contact( "FC4_F+" )
      I_Contact( "ETAPA_101" )
      Coil( "MARCA_VACIAA" )
   END_RUNG
   RUNG wire#powerrail
      Contact( "ETAPA_20" )
   END_RUNG wire#w2
   RUNG wire#powerrail
      Contact( "ETAPA_9" )
      wire#w3
      Contact( "FC5_G-" )
      I_Contact( "ETAPA_101" )
      Move(in := 5.49, out1 => "CILINDRO G")
   END_RUNG
   RUNG wire#powerrail
      Contact( "ETAPA_19" )
   END_RUNG wire#w3
   RUNG wire#powerrail
      Contact( "ETAPA_11" )
      wire#w4
      Contact( "FC6_G+" )
      I_Contact( "ETAPA_101" )
      Move(in := -3.5, out1 => "CILINDRO G")
   END_RUNG
   RUNG wire#powerrail
      Contact( "ETAPA_21" )
   END_RUNG wire#w4
   // the same network as SCL:
   "CILINDRO F" := ("ETAPA_8" OR "ETAPA_18") AND NOT "ETAPA_101";
   "MARCA_VACIAA" := ("ETAPA _10" OR "ETAPA_20") AND "FC4_F+" AND NOT "ETAPA_101";
   IF ("ETAPA_9" OR "ETAPA_19") AND "FC5_G-" AND NOT "ETAPA_101" THEN "CILINDRO G" := 5.49; END_IF;
   IF ("ETAPA_11" OR "ETAPA_21") AND "FC6_G+" AND NOT "ETAPA_101" THEN "CILINDRO G" := -3.5; END_IF;
END_REGION

REGION Network 4: PROGRAMACIÓN IMAGEN DE CONTROL HMI (PROCESO SALIDA)
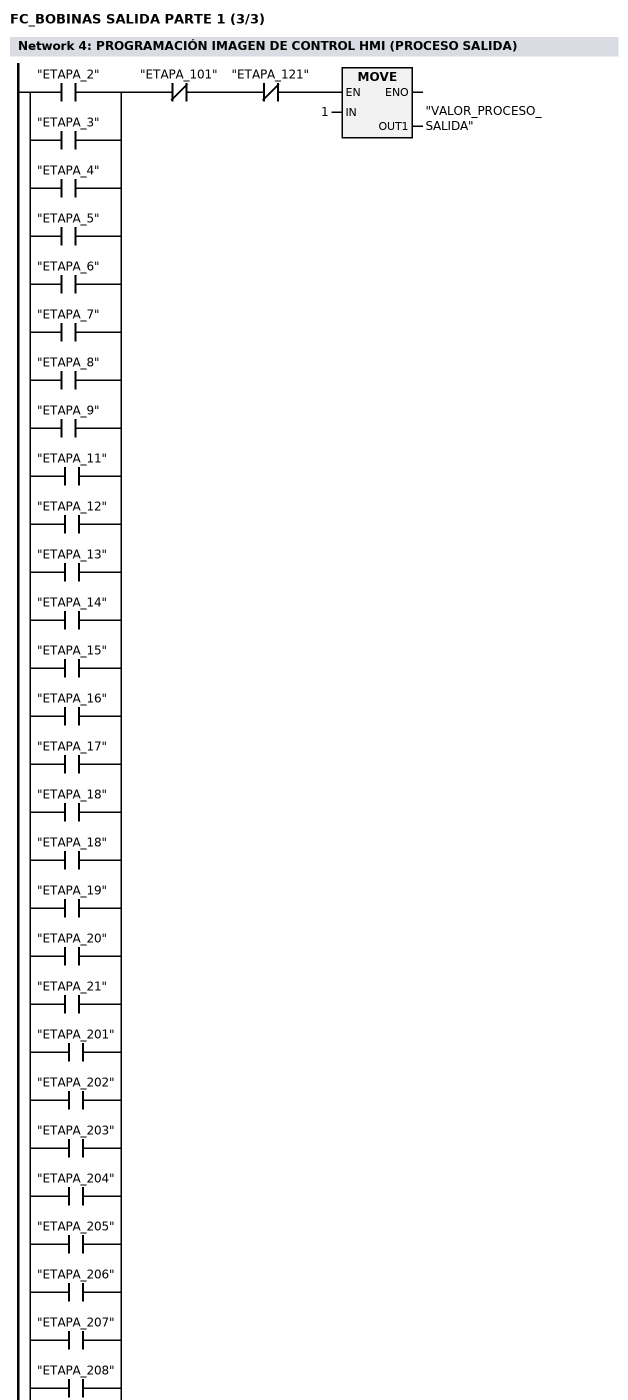
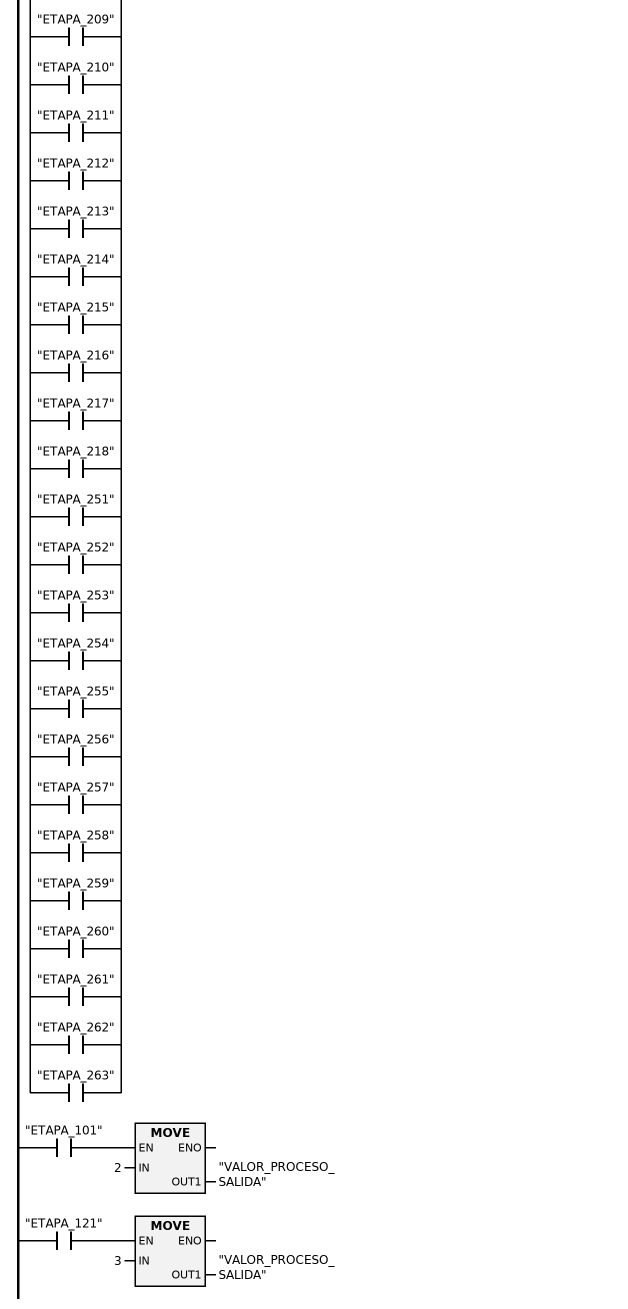
   RUNG wire#powerrail
      Contact( "ETAPA_2" )
      wire#w1
      I_Contact( "ETAPA_101" )
      I_Contact( "ETAPA_121" )
      Move(in := 1, out1 => "VALOR_PROCESO_SALIDA")
   END_RUNG
   RUNG wire#powerrail
      Contact( "ETAPA_3" )
   END_RUNG wire#w1
   RUNG wire#powerrail
      Contact( "ETAPA_4" )
   END_RUNG wire#w1
   RUNG wire#powerrail
      Contact( "ETAPA_5" )
   END_RUNG wire#w1
   RUNG wire#powerrail
      Contact( "ETAPA_6" )
   END_RUNG wire#w1
   RUNG wire#powerrail
      Contact( "ETAPA_7" )
   END_RUNG wire#w1
   RUNG wire#powerrail
      Contact( "ETAPA_8" )
   END_RUNG wire#w1
   RUNG wire#powerrail
      Contact( "ETAPA_9" )
   END_RUNG wire#w1
   RUNG wire#powerrail
      Contact( "ETAPA_11" )
   END_RUNG wire#w1
   RUNG wire#powerrail
      Contact( "ETAPA_12" )
   END_RUNG wire#w1
   RUNG wire#powerrail
      Contact( "ETAPA_13" )
   END_RUNG wire#w1
   RUNG wire#powerrail
      Contact( "ETAPA_14" )
   END_RUNG wire#w1
   RUNG wire#powerrail
      Contact( "ETAPA_15" )
   END_RUNG wire#w1
   RUNG wire#powerrail
      Contact( "ETAPA_16" )
   END_RUNG wire#w1
   RUNG wire#powerrail
      Contact( "ETAPA_17" )
   END_RUNG wire#w1
   RUNG wire#powerrail
      Contact( "ETAPA_18" )
   END_RUNG wire#w1
   RUNG wire#powerrail
      Contact( "ETAPA_18" )
   END_RUNG wire#w1
   RUNG wire#powerrail
      Contact( "ETAPA_19" )
   END_RUNG wire#w1
   RUNG wire#powerrail
      Contact( "ETAPA_20" )
   END_RUNG wire#w1
   RUNG wire#powerrail
      Contact( "ETAPA_21" )
   END_RUNG wire#w1
   RUNG wire#powerrail
      Contact( "ETAPA_201" )
   END_RUNG wire#w1
   RUNG wire#powerrail
      Contact( "ETAPA_202" )
   END_RUNG wire#w1
   RUNG wire#powerrail
      Contact( "ETAPA_203" )
   END_RUNG wire#w1
   RUNG wire#powerrail
      Contact( "ETAPA_204" )
   END_RUNG wire#w1
   RUNG wire#powerrail
      Contact( "ETAPA_205" )
   END_RUNG wire#w1
   RUNG wire#powerrail
      Contact( "ETAPA_206" )
   END_RUNG wire#w1
   RUNG wire#powerrail
      Contact( "ETAPA_207" )
   END_RUNG wire#w1
   RUNG wire#powerrail
      Contact( "ETAPA_208" )
   END_RUNG wire#w1
   RUNG wire#powerrail
      Contact( "ETAPA_209" )
   END_RUNG wire#w1
   RUNG wire#powerrail
      Contact( "ETAPA_210" )
   END_RUNG wire#w1
   RUNG wire#powerrail
      Contact( "ETAPA_211" )
   END_RUNG wire#w1
   RUNG wire#powerrail
      Contact( "ETAPA_212" )
   END_RUNG wire#w1
   RUNG wire#powerrail
      Contact( "ETAPA_213" )
   END_RUNG wire#w1
   RUNG wire#powerrail
      Contact( "ETAPA_214" )
   END_RUNG wire#w1
   RUNG wire#powerrail
      Contact( "ETAPA_215" )
   END_RUNG wire#w1
   RUNG wire#powerrail
      Contact( "ETAPA_216" )
   END_RUNG wire#w1
   RUNG wire#powerrail
      Contact( "ETAPA_217" )
   END_RUNG wire#w1
   RUNG wire#powerrail
      Contact( "ETAPA_218" )
   END_RUNG wire#w1
   RUNG wire#powerrail
      Contact( "ETAPA_251" )
   END_RUNG wire#w1
   RUNG wire#powerrail
      Contact( "ETAPA_252" )
   END_RUNG wire#w1
   RUNG wire#powerrail
      Contact( "ETAPA_253" )
   END_RUNG wire#w1
   RUNG wire#powerrail
      Contact( "ETAPA_254" )
   END_RUNG wire#w1
   RUNG wire#powerrail
      Contact( "ETAPA_255" )
   END_RUNG wire#w1
   RUNG wire#powerrail
      Contact( "ETAPA_256" )
   END_RUNG wire#w1
   RUNG wire#powerrail
      Contact( "ETAPA_257" )
   END_RUNG wire#w1
   RUNG wire#powerrail
      Contact( "ETAPA_258" )
   END_RUNG wire#w1
   RUNG wire#powerrail
      Contact( "ETAPA_259" )
   END_RUNG wire#w1
   RUNG wire#powerrail
      Contact( "ETAPA_260" )
   END_RUNG wire#w1
   RUNG wire#powerrail
      Contact( "ETAPA_261" )
   END_RUNG wire#w1
   RUNG wire#powerrail
      Contact( "ETAPA_262" )
   END_RUNG wire#w1
   RUNG wire#powerrail
      Contact( "ETAPA_263" )
   END_RUNG wire#w1
   RUNG wire#powerrail
      Contact( "ETAPA_101" )
      Move(in := 2, out1 => "VALOR_PROCESO_SALIDA")
   END_RUNG
   RUNG wire#powerrail
      Contact( "ETAPA_121" )
      Move(in := 3, out1 => "VALOR_PROCESO_SALIDA")
   END_RUNG
   // the same network as SCL:
   IF ("ETAPA_2" OR "ETAPA_3" OR "ETAPA_4" OR "ETAPA_5" OR "ETAPA_6" OR "ETAPA_7" OR "ETAPA_8" OR "ETAPA_9" OR "ETAPA_11" OR "ETAPA_12" OR "ETAPA_13" OR "ETAPA_14" OR "ETAPA_15" OR "ETAPA_16" OR "ETAPA_17" OR "ETAPA_18" OR "ETAPA_18" OR "ETAPA_19" OR "ETAPA_20" OR "ETAPA_21" OR "ETAPA_201" OR "ETAPA_202" OR "ETAPA_203" OR "ETAPA_204" OR "ETAPA_205" OR "ETAPA_206" OR "ETAPA_207" OR "ETAPA_208" OR "ETAPA_209" OR "ETAPA_210" OR "ETAPA_211" OR "ETAPA_212" OR "ETAPA_213" OR "ETAPA_214" OR "ETAPA_215" OR "ETAPA_216" OR "ETAPA_217" OR "ETAPA_218" OR "ETAPA_251" OR "ETAPA_252" OR "ETAPA_253" OR "ETAPA_254" OR "ETAPA_255" OR "ETAPA_256" OR "ETAPA_257" OR "ETAPA_258" OR "ETAPA_259" OR "ETAPA_260" OR "ETAPA_261" OR "ETAPA_262" OR "ETAPA_263") AND NOT "ETAPA_101" AND NOT "ETAPA_121" THEN
       "VALOR_PROCESO_SALIDA" := 1;
   END_IF;
   IF "ETAPA_101" THEN "VALOR_PROCESO_SALIDA" := 2; END_IF;
   IF "ETAPA_121" THEN "VALOR_PROCESO_SALIDA" := 3; END_IF;
END_REGION
END_FUNCTION

FUNCTION "FC_PARADA SALIDA" : Void   // FC3, LAD
{ S7_Optimized_Access := 'TRUE' }
VERSION : 0.1
// EN ESTE BLOQUE SE MUESTRA LA PARADA DEL PROCESO DE SALIDA
   VAR_TEMP   // added for the SCL form of the ladder/FBD networks
      _w1 : Bool;
   END_VAR
BEGIN

REGION Network 1: PROGRAMACIÓN DE LA PARADA POR PULSADOR DE PARO
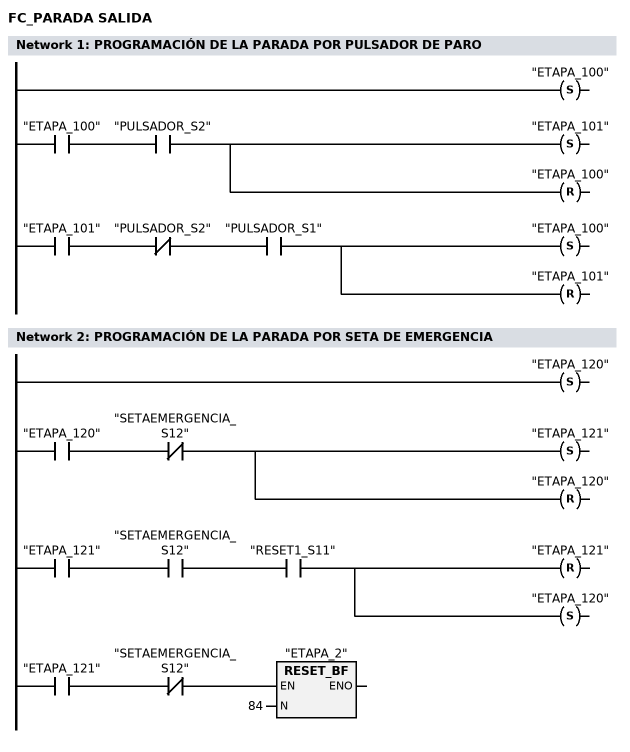
   RUNG wire#powerrail
      S_Coil( "ETAPA_100" )
   END_RUNG
   RUNG wire#powerrail
      Contact( "ETAPA_100" )
      Contact( "PULSADOR_S2" )
      wire#w1
      S_Coil( "ETAPA_101" )
   END_RUNG
   RUNG wire#w1
      R_Coil( "ETAPA_100" )
   END_RUNG
   RUNG wire#powerrail
      Contact( "ETAPA_101" )
      I_Contact( "PULSADOR_S2" )
      Contact( "PULSADOR_S1" )
      wire#w2
      S_Coil( "ETAPA_100" )
   END_RUNG
   RUNG wire#w2
      R_Coil( "ETAPA_101" )
   END_RUNG
   // the same network as SCL:
   "ETAPA_100" := TRUE;
   IF "ETAPA_100" AND "PULSADOR_S2" THEN
       "ETAPA_101" := TRUE;
       "ETAPA_100" := FALSE;
   END_IF;
   IF "ETAPA_101" AND NOT "PULSADOR_S2" AND "PULSADOR_S1" THEN
       "ETAPA_100" := TRUE;
       "ETAPA_101" := FALSE;
   END_IF;
END_REGION

REGION Network 2: PROGRAMACIÓN DE LA PARADA POR SETA DE EMERGENCIA
   // no SCL statement known for RBitfield: written as a call
   "ETAPA_120" := TRUE;
   IF "ETAPA_120" AND NOT "SETAEMERGENCIA_S12" THEN
       "ETAPA_121" := TRUE;
       "ETAPA_120" := FALSE;
   END_IF;
   #_w1 := "ETAPA_121" AND "SETAEMERGENCIA_S12" AND "RESET1_S11";
   IF #_w1 THEN
       "ETAPA_121" := FALSE;
       "ETAPA_120" := TRUE;
   END_IF;
   IF "ETAPA_121" AND NOT "SETAEMERGENCIA_S12" THEN RESET_BF(operand := "ETAPA_2", n := 84); END_IF;
END_REGION
END_FUNCTION

FUNCTION "FC_SECUENCIA ENTRADA" : Void   // FC4, LAD
{ S7_Optimized_Access := 'TRUE' }
VERSION : 0.1
// EN ESTE BLOQUE SE ENCUENTRA LA PROGRAMACIÓN DE LA SECUENCIA DEL PROCESO DE ENTRADA, DESDE EL PRINCIPIO DEL PROCESO HASTA  QUE LLEGA A LA ENTRADA DEL ROBOT
   VAR_TEMP   // added for the SCL form of the ladder/FBD networks
      _w1 : Bool;
   END_VAR
BEGIN

REGION Network 1: SET DE LA ETAPA 0
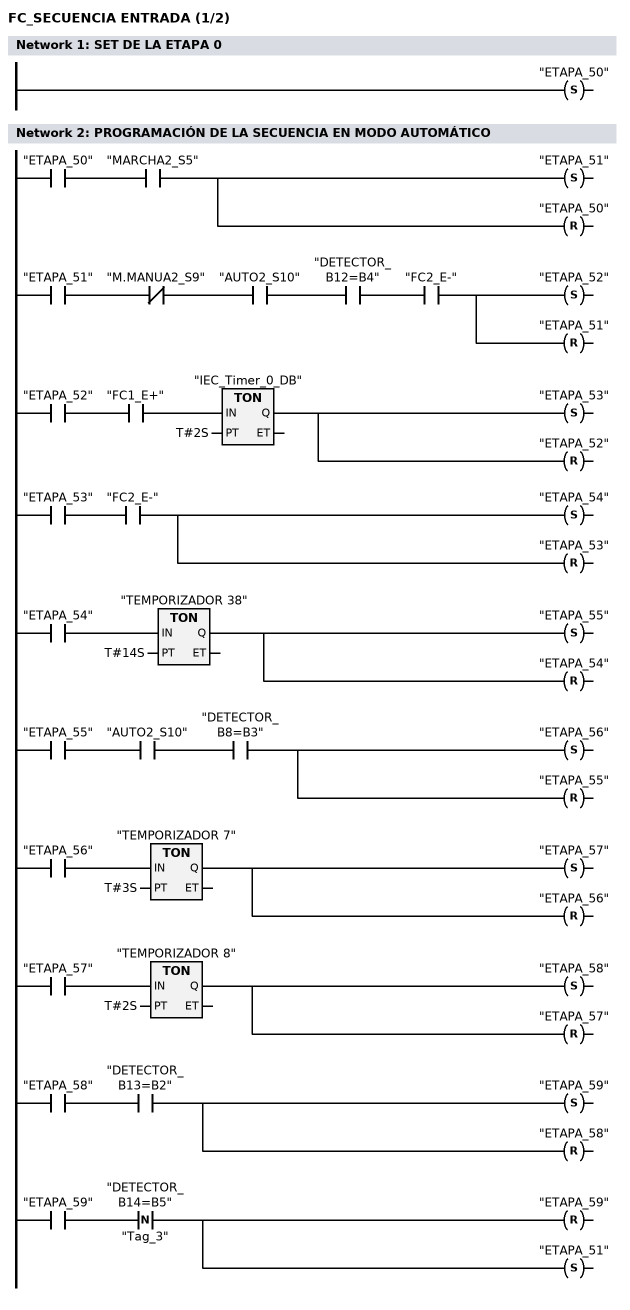
   RUNG wire#powerrail
      S_Coil( "ETAPA_50" )
   END_RUNG
   // the same network as SCL:
   "ETAPA_50" := TRUE;
END_REGION

REGION Network 2: PROGRAMACIÓN DE LA SECUENCIA EN MODO AUTOMÁTICO
   IF "ETAPA_50" AND "MARCHA2_S5" THEN
       "ETAPA_51" := TRUE;
       "ETAPA_50" := FALSE;
   END_IF;
   IF "ETAPA_51" AND NOT "M.MANUA2_S9" AND "AUTO2_S10" AND "DETECTOR_B12=B4" AND "FC2_E-" THEN
       "ETAPA_52" := TRUE;
       "ETAPA_51" := FALSE;
   END_IF;
   "IEC_Timer_0_DB".TON(IN := "ETAPA_52" AND "FC1_E+", PT := T#2S);
   IF "IEC_Timer_0_DB".Q THEN
       "ETAPA_53" := TRUE;
       "ETAPA_52" := FALSE;
   END_IF;
   IF "ETAPA_53" AND "FC2_E-" THEN
       "ETAPA_54" := TRUE;
       "ETAPA_53" := FALSE;
   END_IF;
   "TEMPORIZADOR 38".TON(IN := "ETAPA_54", PT := T#14S);
   IF "TEMPORIZADOR 38".Q THEN
       "ETAPA_55" := TRUE;
       "ETAPA_54" := FALSE;
   END_IF;
   IF "ETAPA_55" AND "AUTO2_S10" AND "DETECTOR_B8=B3" THEN
       "ETAPA_56" := TRUE;
       "ETAPA_55" := FALSE;
   END_IF;
   "TEMPORIZADOR 7".TON(IN := "ETAPA_56", PT := T#3S);
   IF "TEMPORIZADOR 7".Q THEN
       "ETAPA_57" := TRUE;
       "ETAPA_56" := FALSE;
   END_IF;
   "TEMPORIZADOR 8".TON(IN := "ETAPA_57", PT := T#2S);
   IF "TEMPORIZADOR 8".Q THEN
       "ETAPA_58" := TRUE;
       "ETAPA_57" := FALSE;
   END_IF;
   IF "ETAPA_58" AND "DETECTOR_B13=B2" THEN
       "ETAPA_59" := TRUE;
       "ETAPA_58" := FALSE;
   END_IF;
   #_w1 := "ETAPA_59" AND NOT "DETECTOR_B14=B5" AND "Tag_3";   // falling edge of "DETECTOR_B14=B5"
   "Tag_3" := "DETECTOR_B14=B5";
   IF #_w1 THEN
       "ETAPA_59" := FALSE;
       "ETAPA_51" := TRUE;
   END_IF;
END_REGION

REGION Network 3: PROGRAMACIÓN DE LA SECUENCIA EN MODO MANUAL
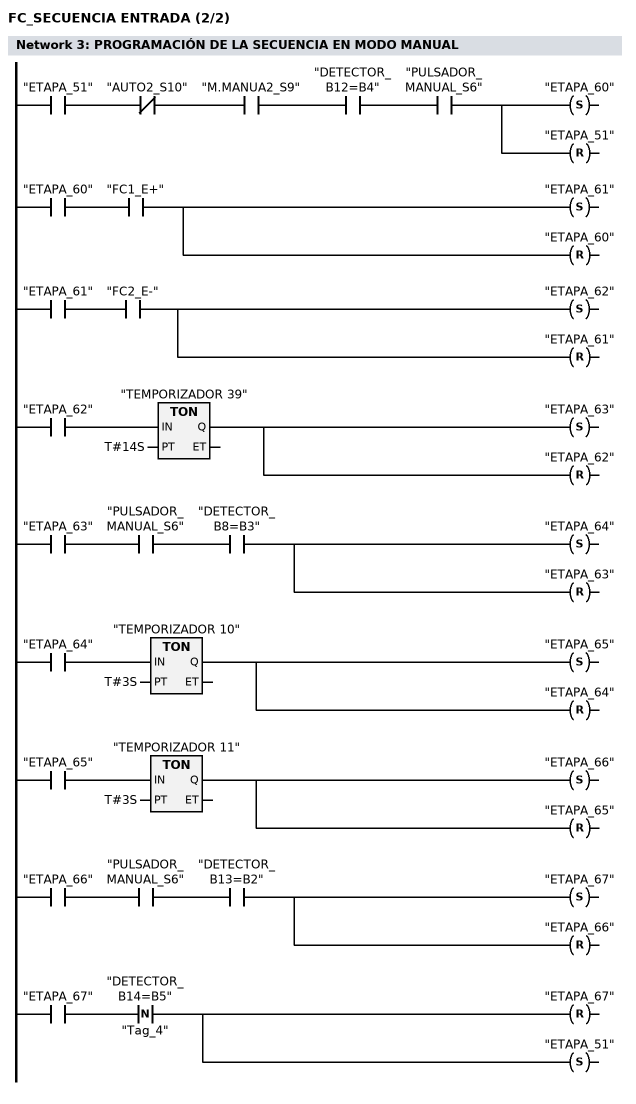
   IF "ETAPA_51" AND NOT "AUTO2_S10" AND "M.MANUA2_S9" AND "DETECTOR_B12=B4" AND "PULSADOR_MANUAL_S6" THEN
       "ETAPA_60" := TRUE;
       "ETAPA_51" := FALSE;
   END_IF;
   IF "ETAPA_60" AND "FC1_E+" THEN
       "ETAPA_61" := TRUE;
       "ETAPA_60" := FALSE;
   END_IF;
   IF "ETAPA_61" AND "FC2_E-" THEN
       "ETAPA_62" := TRUE;
       "ETAPA_61" := FALSE;
   END_IF;
   "TEMPORIZADOR 39".TON(IN := "ETAPA_62", PT := T#14S);
   IF "TEMPORIZADOR 39".Q THEN
       "ETAPA_63" := TRUE;
       "ETAPA_62" := FALSE;
   END_IF;
   IF "ETAPA_63" AND "PULSADOR_MANUAL_S6" AND "DETECTOR_B8=B3" THEN
       "ETAPA_64" := TRUE;
       "ETAPA_63" := FALSE;
   END_IF;
   "TEMPORIZADOR 10".TON(IN := "ETAPA_64", PT := T#3S);
   IF "TEMPORIZADOR 10".Q THEN
       "ETAPA_65" := TRUE;
       "ETAPA_64" := FALSE;
   END_IF;
   "TEMPORIZADOR 11".TON(IN := "ETAPA_65", PT := T#3S);
   IF "TEMPORIZADOR 11".Q THEN
       "ETAPA_66" := TRUE;
       "ETAPA_65" := FALSE;
   END_IF;
   IF "ETAPA_66" AND "PULSADOR_MANUAL_S6" AND "DETECTOR_B13=B2" THEN
       "ETAPA_67" := TRUE;
       "ETAPA_66" := FALSE;
   END_IF;
   #_w1 := "ETAPA_67" AND NOT "DETECTOR_B14=B5" AND "Tag_4";   // falling edge of "DETECTOR_B14=B5"
   "Tag_4" := "DETECTOR_B14=B5";
   IF #_w1 THEN
       "ETAPA_67" := FALSE;
       "ETAPA_51" := TRUE;
   END_IF;
END_REGION
END_FUNCTION

FUNCTION "FC_BOBINAS ENTRADA" : Void   // FC5, LAD
{ S7_Optimized_Access := 'TRUE' }
VERSION : 0.1
// EN ESTE BLOQUE SE ENCUENTRA LA ASIGNACIÓN DE CADA ETAPA CON EL ACTUADOR QUE CORRESPONDE, DESDE EL PRINCIPIO DEL PROCESO HASTA  QUE LLEGA A LA ENTRADA DEL ROBOT
BEGIN

REGION Network 1: ASIGNACIÓN DE CADA BOBINA CON SU CORRESPONDIENTE ACTUADOR; PROCESO DE ENTRADA
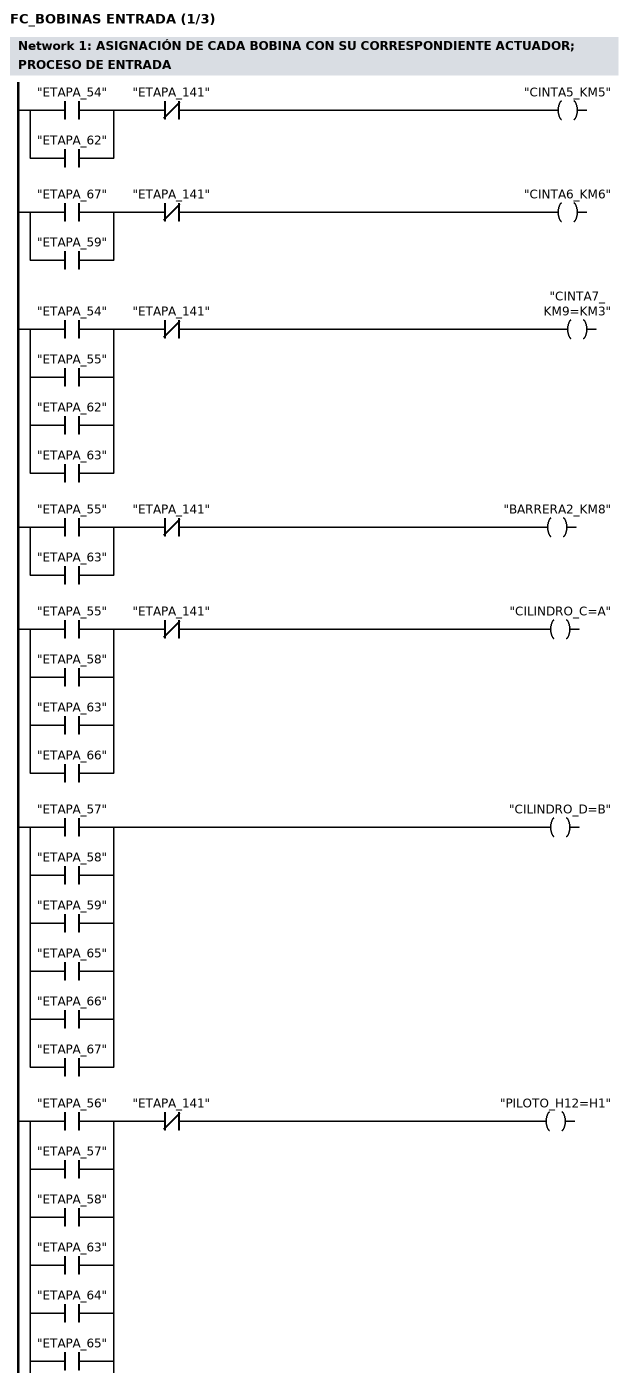
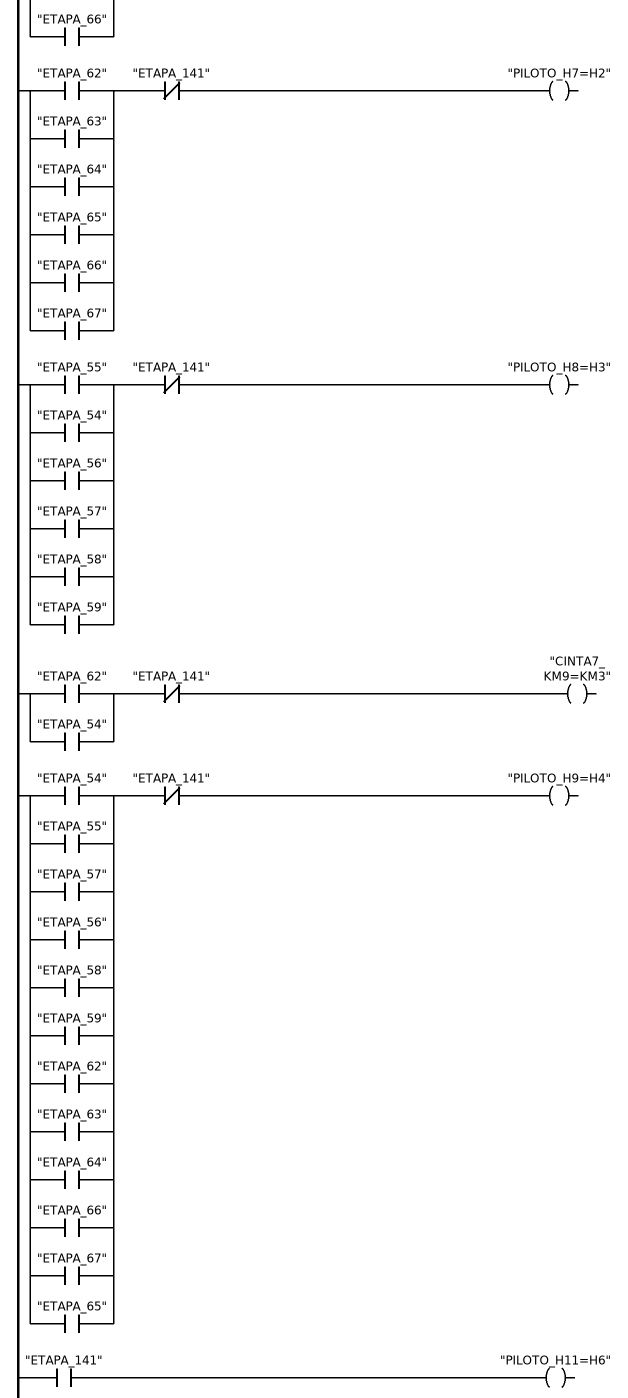
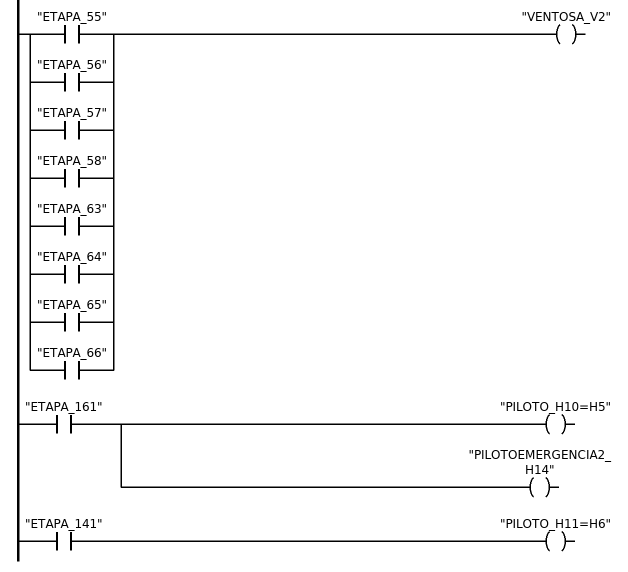
   RUNG wire#powerrail
      Contact( "ETAPA_54" )
      wire#w1
      I_Contact( "ETAPA_141" )
      Coil( "CINTA5_KM5" )
   END_RUNG
   RUNG wire#powerrail
      Contact( "ETAPA_62" )
   END_RUNG wire#w1
   RUNG wire#powerrail
      Contact( "ETAPA_67" )
      wire#w2
      I_Contact( "ETAPA_141" )
      Coil( "CINTA6_KM6" )
   END_RUNG
   RUNG wire#powerrail
      Contact( "ETAPA_59" )
   END_RUNG wire#w2
   RUNG wire#powerrail
      Contact( "ETAPA_54" )
      wire#w3
      I_Contact( "ETAPA_141" )
      Coil( "CINTA7_KM9=KM3" )
   END_RUNG
   RUNG wire#powerrail
      Contact( "ETAPA_55" )
   END_RUNG wire#w3
   RUNG wire#powerrail
      Contact( "ETAPA_62" )
   END_RUNG wire#w3
   RUNG wire#powerrail
      Contact( "ETAPA_63" )
   END_RUNG wire#w3
   RUNG wire#powerrail
      Contact( "ETAPA_55" )
      wire#w4
      I_Contact( "ETAPA_141" )
      Coil( "BARRERA2_KM8" )
   END_RUNG
   RUNG wire#powerrail
      Contact( "ETAPA_63" )
   END_RUNG wire#w4
   RUNG wire#powerrail
      Contact( "ETAPA_55" )
      wire#w5
      I_Contact( "ETAPA_141" )
      Coil( "CILINDRO_C=A" )
   END_RUNG
   RUNG wire#powerrail
      Contact( "ETAPA_58" )
   END_RUNG wire#w5
   RUNG wire#powerrail
      Contact( "ETAPA_63" )
   END_RUNG wire#w5
   RUNG wire#powerrail
      Contact( "ETAPA_66" )
   END_RUNG wire#w5
   RUNG wire#powerrail
      Contact( "ETAPA_57" )
      wire#w6
      Coil( "CILINDRO_D=B" )
   END_RUNG
   RUNG wire#powerrail
      Contact( "ETAPA_58" )
   END_RUNG wire#w6
   RUNG wire#powerrail
      Contact( "ETAPA_59" )
   END_RUNG wire#w6
   RUNG wire#powerrail
      Contact( "ETAPA_65" )
   END_RUNG wire#w6
   RUNG wire#powerrail
      Contact( "ETAPA_66" )
   END_RUNG wire#w6
   RUNG wire#powerrail
      Contact( "ETAPA_67" )
   END_RUNG wire#w6
   RUNG wire#powerrail
      Contact( "ETAPA_56" )
      wire#w7
      I_Contact( "ETAPA_141" )
      Coil( "PILOTO_H12=H1" )
   END_RUNG
   RUNG wire#powerrail
      Contact( "ETAPA_57" )
   END_RUNG wire#w7
   RUNG wire#powerrail
      Contact( "ETAPA_58" )
   END_RUNG wire#w7
   RUNG wire#powerrail
      Contact( "ETAPA_63" )
   END_RUNG wire#w7
   RUNG wire#powerrail
      Contact( "ETAPA_64" )
   END_RUNG wire#w7
   RUNG wire#powerrail
      Contact( "ETAPA_65" )
   END_RUNG wire#w7
   RUNG wire#powerrail
      Contact( "ETAPA_66" )
   END_RUNG wire#w7
   RUNG wire#powerrail
      Contact( "ETAPA_62" )
      wire#w8
      I_Contact( "ETAPA_141" )
      Coil( "PILOTO_H7=H2" )
   END_RUNG
   RUNG wire#powerrail
      Contact( "ETAPA_63" )
   END_RUNG wire#w8
   RUNG wire#powerrail
      Contact( "ETAPA_64" )
   END_RUNG wire#w8
   RUNG wire#powerrail
      Contact( "ETAPA_65" )
   END_RUNG wire#w8
   RUNG wire#powerrail
      Contact( "ETAPA_66" )
   END_RUNG wire#w8
   RUNG wire#powerrail
      Contact( "ETAPA_67" )
   END_RUNG wire#w8
   RUNG wire#powerrail
      Contact( "ETAPA_55" )
      wire#w9
      I_Contact( "ETAPA_141" )
      Coil( "PILOTO_H8=H3" )
   END_RUNG
   RUNG wire#powerrail
      Contact( "ETAPA_54" )
   END_RUNG wire#w9
   RUNG wire#powerrail
      Contact( "ETAPA_56" )
   END_RUNG wire#w9
   RUNG wire#powerrail
      Contact( "ETAPA_57" )
   END_RUNG wire#w9
   RUNG wire#powerrail
      Contact( "ETAPA_58" )
   END_RUNG wire#w9
   RUNG wire#powerrail
      Contact( "ETAPA_59" )
   END_RUNG wire#w9
   RUNG wire#powerrail
      Contact( "ETAPA_62" )
      wire#w10
      I_Contact( "ETAPA_141" )
      Coil( "CINTA7_KM9=KM3" )
   END_RUNG
   RUNG wire#powerrail
      Contact( "ETAPA_54" )
   END_RUNG wire#w10
   RUNG wire#powerrail
      Contact( "ETAPA_54" )
      wire#w11
      I_Contact( "ETAPA_141" )
      Coil( "PILOTO_H9=H4" )
   END_RUNG
   RUNG wire#powerrail
      Contact( "ETAPA_55" )
   END_RUNG wire#w11
   RUNG wire#powerrail
      Contact( "ETAPA_57" )
   END_RUNG wire#w11
   RUNG wire#powerrail
      Contact( "ETAPA_56" )
   END_RUNG wire#w11
   RUNG wire#powerrail
      Contact( "ETAPA_58" )
   END_RUNG wire#w11
   RUNG wire#powerrail
      Contact( "ETAPA_59" )
   END_RUNG wire#w11
   RUNG wire#powerrail
      Contact( "ETAPA_62" )
   END_RUNG wire#w11
   RUNG wire#powerrail
      Contact( "ETAPA_63" )
   END_RUNG wire#w11
   RUNG wire#powerrail
      Contact( "ETAPA_64" )
   END_RUNG wire#w11
   RUNG wire#powerrail
      Contact( "ETAPA_66" )
   END_RUNG wire#w11
   RUNG wire#powerrail
      Contact( "ETAPA_67" )
   END_RUNG wire#w11
   RUNG wire#powerrail
      Contact( "ETAPA_65" )
   END_RUNG wire#w11
   RUNG wire#powerrail
      Contact( "ETAPA_141" )
      Coil( "PILOTO_H11=H6" )
   END_RUNG
   RUNG wire#powerrail
      Contact( "ETAPA_55" )
      wire#w12
      Coil( "VENTOSA_V2" )
   END_RUNG
   RUNG wire#powerrail
      Contact( "ETAPA_56" )
   END_RUNG wire#w12
   RUNG wire#powerrail
      Contact( "ETAPA_57" )
   END_RUNG wire#w12
   RUNG wire#powerrail
      Contact( "ETAPA_58" )
   END_RUNG wire#w12
   RUNG wire#powerrail
      Contact( "ETAPA_63" )
   END_RUNG wire#w12
   RUNG wire#powerrail
      Contact( "ETAPA_64" )
   END_RUNG wire#w12
   RUNG wire#powerrail
      Contact( "ETAPA_65" )
   END_RUNG wire#w12
   RUNG wire#powerrail
      Contact( "ETAPA_66" )
   END_RUNG wire#w12
   RUNG wire#powerrail
      Contact( "ETAPA_161" )
      wire#w13
      Coil( "PILOTO_H10=H5" )
   END_RUNG
   RUNG wire#w13
      Coil( "PILOTOEMERGENCIA2_H14" )
   END_RUNG
   RUNG wire#powerrail
      Contact( "ETAPA_141" )
      Coil( "PILOTO_H11=H6" )
   END_RUNG
   // the same network as SCL:
   "CINTA5_KM5" := ("ETAPA_54" OR "ETAPA_62") AND NOT "ETAPA_141";
   "CINTA6_KM6" := ("ETAPA_67" OR "ETAPA_59") AND NOT "ETAPA_141";
   "CINTA7_KM9=KM3" := ("ETAPA_54" OR "ETAPA_55" OR "ETAPA_62" OR "ETAPA_63") AND NOT "ETAPA_141";
   "BARRERA2_KM8" := ("ETAPA_55" OR "ETAPA_63") AND NOT "ETAPA_141";
   "CILINDRO_C=A" := ("ETAPA_55" OR "ETAPA_58" OR "ETAPA_63" OR "ETAPA_66") AND NOT "ETAPA_141";
   "CILINDRO_D=B" := "ETAPA_57" OR "ETAPA_58" OR "ETAPA_59" OR "ETAPA_65" OR "ETAPA_66" OR "ETAPA_67";
   "PILOTO_H12=H1" := ("ETAPA_56" OR "ETAPA_57" OR "ETAPA_58" OR "ETAPA_63" OR "ETAPA_64" OR "ETAPA_65" OR "ETAPA_66") AND NOT "ETAPA_141";
   "PILOTO_H7=H2" := ("ETAPA_62" OR "ETAPA_63" OR "ETAPA_64" OR "ETAPA_65" OR "ETAPA_66" OR "ETAPA_67") AND NOT "ETAPA_141";
   "PILOTO_H8=H3" := ("ETAPA_55" OR "ETAPA_54" OR "ETAPA_56" OR "ETAPA_57" OR "ETAPA_58" OR "ETAPA_59") AND NOT "ETAPA_141";
   "CINTA7_KM9=KM3" := ("ETAPA_62" OR "ETAPA_54") AND NOT "ETAPA_141";
   "PILOTO_H9=H4" := ("ETAPA_54" OR "ETAPA_55" OR "ETAPA_57" OR "ETAPA_56" OR "ETAPA_58" OR "ETAPA_59" OR "ETAPA_62" OR "ETAPA_63" OR "ETAPA_64" OR "ETAPA_66" OR "ETAPA_67" OR "ETAPA_65") AND NOT "ETAPA_141";
   "PILOTO_H11=H6" := "ETAPA_141";
   "VENTOSA_V2" := "ETAPA_55" OR "ETAPA_56" OR "ETAPA_57" OR "ETAPA_58" OR "ETAPA_63" OR "ETAPA_64" OR "ETAPA_65" OR "ETAPA_66";
   "PILOTO_H10=H5" := "ETAPA_161";
   "PILOTOEMERGENCIA2_H14" := "ETAPA_161";
   "PILOTO_H11=H6" := "ETAPA_141";
END_REGION

REGION Network 2: ASIGNACIÓN Y PROGRAMACIÓN CILINDRO E
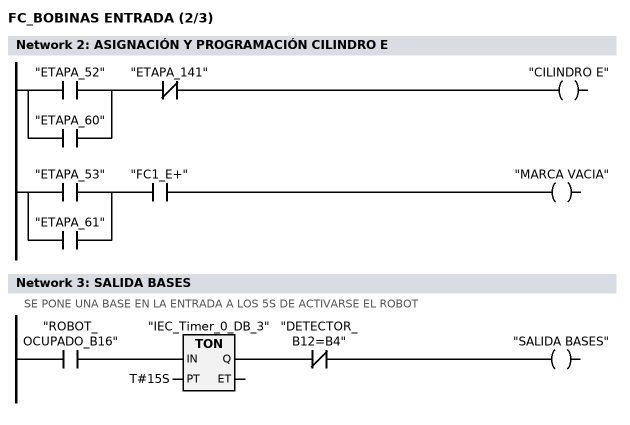
   RUNG wire#powerrail
      Contact( "ETAPA_52" )
      wire#w1
      I_Contact( "ETAPA_141" )
      Coil( "CILINDRO E" )
   END_RUNG
   RUNG wire#powerrail
      Contact( "ETAPA_60" )
   END_RUNG wire#w1
   RUNG wire#powerrail
      Contact( "ETAPA_53" )
      wire#w2
      Contact( "FC1_E+" )
      Coil( "MARCA VACIA" )
   END_RUNG
   RUNG wire#powerrail
      Contact( "ETAPA_61" )
   END_RUNG wire#w2
   // the same network as SCL:
   "CILINDRO E" := ("ETAPA_52" OR "ETAPA_60") AND NOT "ETAPA_141";
   "MARCA VACIA" := ("ETAPA_53" OR "ETAPA_61") AND "FC1_E+";
END_REGION

REGION Network 3: SALIDA BASES
   // SE PONE UNA BASE EN LA ENTRADA A LOS 5S DE ACTIVARSE EL ROBOT
   "IEC_Timer_0_DB_3".TON(IN := "ROBOT_OCUPADO_B16", PT := T#15S);
   "SALIDA BASES" := "IEC_Timer_0_DB_3".Q AND NOT "DETECTOR_B12=B4";
END_REGION

REGION Network 4: PROGRAMACIÓN IMAGEN DE CONTROL HMI (PROCESO ENTRADA)
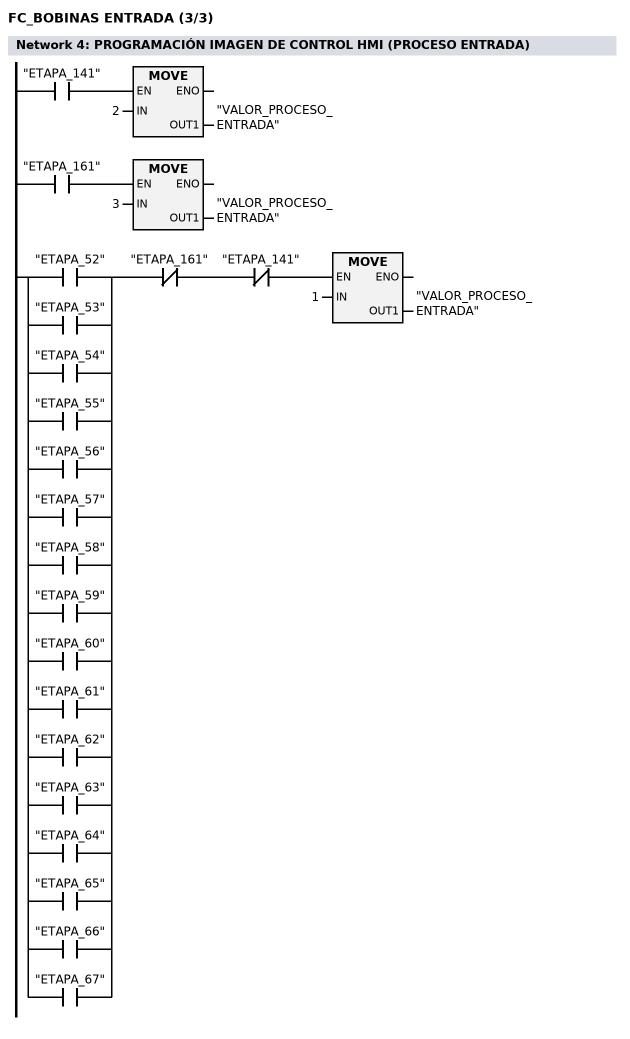
   RUNG wire#powerrail
      Contact( "ETAPA_141" )
      Move(in := 2, out1 => "VALOR_PROCESO_ENTRADA")
   END_RUNG
   RUNG wire#powerrail
      Contact( "ETAPA_161" )
      Move(in := 3, out1 => "VALOR_PROCESO_ENTRADA")
   END_RUNG
   RUNG wire#powerrail
      Contact( "ETAPA_52" )
      wire#w1
      I_Contact( "ETAPA_161" )
      I_Contact( "ETAPA_141" )
      Move(in := 1, out1 => "VALOR_PROCESO_ENTRADA")
   END_RUNG
   RUNG wire#powerrail
      Contact( "ETAPA_53" )
   END_RUNG wire#w1
   RUNG wire#powerrail
      Contact( "ETAPA_54" )
   END_RUNG wire#w1
   RUNG wire#powerrail
      Contact( "ETAPA_55" )
   END_RUNG wire#w1
   RUNG wire#powerrail
      Contact( "ETAPA_56" )
   END_RUNG wire#w1
   RUNG wire#powerrail
      Contact( "ETAPA_57" )
   END_RUNG wire#w1
   RUNG wire#powerrail
      Contact( "ETAPA_58" )
   END_RUNG wire#w1
   RUNG wire#powerrail
      Contact( "ETAPA_59" )
   END_RUNG wire#w1
   RUNG wire#powerrail
      Contact( "ETAPA_60" )
   END_RUNG wire#w1
   RUNG wire#powerrail
      Contact( "ETAPA_61" )
   END_RUNG wire#w1
   RUNG wire#powerrail
      Contact( "ETAPA_62" )
   END_RUNG wire#w1
   RUNG wire#powerrail
      Contact( "ETAPA_63" )
   END_RUNG wire#w1
   RUNG wire#powerrail
      Contact( "ETAPA_64" )
   END_RUNG wire#w1
   RUNG wire#powerrail
      Contact( "ETAPA_65" )
   END_RUNG wire#w1
   RUNG wire#powerrail
      Contact( "ETAPA_66" )
   END_RUNG wire#w1
   RUNG wire#powerrail
      Contact( "ETAPA_67" )
   END_RUNG wire#w1
   // the same network as SCL:
   IF "ETAPA_141" THEN "VALOR_PROCESO_ENTRADA" := 2; END_IF;
   IF "ETAPA_161" THEN "VALOR_PROCESO_ENTRADA" := 3; END_IF;
   IF ("ETAPA_52" OR "ETAPA_53" OR "ETAPA_54" OR "ETAPA_55" OR "ETAPA_56" OR "ETAPA_57" OR "ETAPA_58" OR "ETAPA_59" OR "ETAPA_60" OR "ETAPA_61" OR "ETAPA_62" OR "ETAPA_63" OR "ETAPA_64" OR "ETAPA_65" OR "ETAPA_66" OR "ETAPA_67") AND NOT "ETAPA_161" AND NOT "ETAPA_141" THEN
       "VALOR_PROCESO_ENTRADA" := 1;
   END_IF;
END_REGION
END_FUNCTION

FUNCTION "FC_PARADA ENTRADA" : Void   // FC6, LAD
{ S7_Optimized_Access := 'TRUE' }
VERSION : 0.1
// EN ESTE BLOQUE SE MUESTRA LA PARADA DEL PROCESO DE ENTRADA
   VAR_TEMP   // added for the SCL form of the ladder/FBD networks
      _w1 : Bool;
   END_VAR
BEGIN

REGION Network 1: PARADA DEL PROCESO POR PULSADOR DE PARO
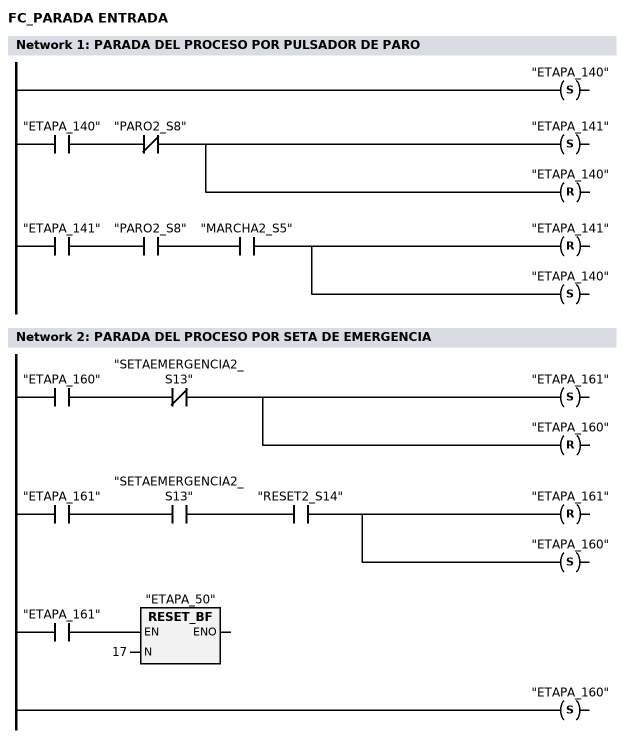
   RUNG wire#powerrail
      S_Coil( "ETAPA_140" )
   END_RUNG
   RUNG wire#powerrail
      Contact( "ETAPA_140" )
      I_Contact( "PARO2_S8" )
      wire#w1
      S_Coil( "ETAPA_141" )
   END_RUNG
   RUNG wire#w1
      R_Coil( "ETAPA_140" )
   END_RUNG
   RUNG wire#powerrail
      Contact( "ETAPA_141" )
      Contact( "PARO2_S8" )
      Contact( "MARCHA2_S5" )
      wire#w2
      R_Coil( "ETAPA_141" )
   END_RUNG
   RUNG wire#w2
      S_Coil( "ETAPA_140" )
   END_RUNG
   // the same network as SCL:
   "ETAPA_140" := TRUE;
   IF "ETAPA_140" AND NOT "PARO2_S8" THEN
       "ETAPA_141" := TRUE;
       "ETAPA_140" := FALSE;
   END_IF;
   #_w1 := "ETAPA_141" AND "PARO2_S8" AND "MARCHA2_S5";
   IF #_w1 THEN
       "ETAPA_141" := FALSE;
       "ETAPA_140" := TRUE;
   END_IF;
END_REGION

REGION Network 2: PARADA DEL PROCESO POR SETA DE EMERGENCIA
   // no SCL statement known for RBitfield: written as a call
   IF "ETAPA_160" AND NOT "SETAEMERGENCIA2_S13" THEN
       "ETAPA_161" := TRUE;
       "ETAPA_160" := FALSE;
   END_IF;
   #_w1 := "ETAPA_161" AND "SETAEMERGENCIA2_S13" AND "RESET2_S14";
   IF #_w1 THEN
       "ETAPA_161" := FALSE;
       "ETAPA_160" := TRUE;
   END_IF;
   IF "ETAPA_161" THEN RESET_BF(operand := "ETAPA_50", n := 17); END_IF;
   "ETAPA_160" := TRUE;
END_REGION
END_FUNCTION

FUNCTION "FC_SECUENCIAROBOT" : Void   // FC7, LAD
{ S7_Optimized_Access := 'TRUE' }
VERSION : 0.1
BEGIN

REGION Network 1
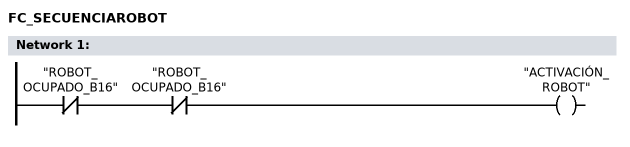
   RUNG wire#powerrail
      I_Contact( "ROBOT_OCUPADO_B16" )
      I_Contact( "ROBOT_OCUPADO_B16" )
      Coil( "ACTIVACIÓN_ROBOT" )
   END_RUNG
   // the same network as SCL:
   "ACTIVACIÓN_ROBOT" := NOT "ROBOT_OCUPADO_B16" AND NOT "ROBOT_OCUPADO_B16";
END_REGION
END_FUNCTION

FUNCTION "FC_SECUENCIA SALIDA PARTE 2_AZUL" : Void   // FC8, LAD
{ S7_Optimized_Access := 'TRUE' }
VERSION : 0.1
// EN ESTE BLOQUE SE ENCUENTRA LA PROGRAMACIÓN DE LA SECUENCIA DESDE QUE LAS CÁMARAS DE VISION DE COLORES DISCRIMAN LA PIEZA AZUL HASTA QUE LA PICK&PLACE XYZ LAS DEJA EN UN PALET
BEGIN

REGION Network 1: SECUENCIA DE SALIDA A PARTIR DE QUE LAS CÁMARAS DISCRIMINAN(CAMINO BASE AZUL)
   // HASTA QUE LA PICK AND PLACE XYZ DEJA LA BASE AZUL EN EL PALET
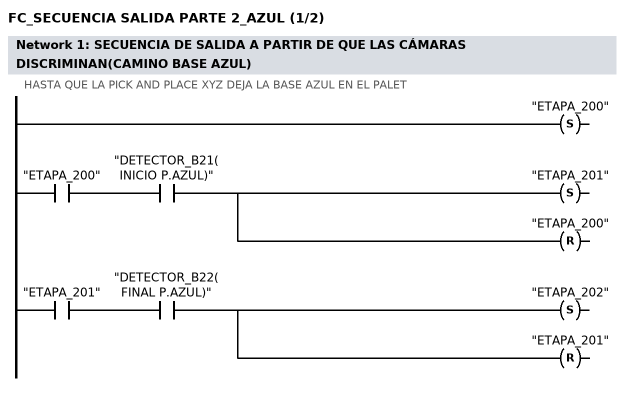
   RUNG wire#powerrail
      S_Coil( "ETAPA_200" )
   END_RUNG
   RUNG wire#powerrail
      Contact( "ETAPA_200" )
      Contact( "DETECTOR_B21(INICIO P.AZUL)" )
      wire#w1
      S_Coil( "ETAPA_201" )
   END_RUNG
   RUNG wire#w1
      R_Coil( "ETAPA_200" )
   END_RUNG
   RUNG wire#powerrail
      Contact( "ETAPA_201" )
      Contact( "DETECTOR_B22(FINAL P.AZUL)" )
      wire#w2
      S_Coil( "ETAPA_202" )
   END_RUNG
   RUNG wire#w2
      R_Coil( "ETAPA_201" )
   END_RUNG
   // the same network as SCL:
   "ETAPA_200" := TRUE;
   IF "ETAPA_200" AND "DETECTOR_B21(INICIO P.AZUL)" THEN
       "ETAPA_201" := TRUE;
       "ETAPA_200" := FALSE;
   END_IF;
   IF "ETAPA_201" AND "DETECTOR_B22(FINAL P.AZUL)" THEN
       "ETAPA_202" := TRUE;
       "ETAPA_201" := FALSE;
   END_IF;
END_REGION

REGION Network 2: SECUENCIA DESDE QUE LLEGA A LA PICK AND PLACE XYZ (BASE AZUL)
   // HASTA QUE LA PIEZA CAE EN EL PALET
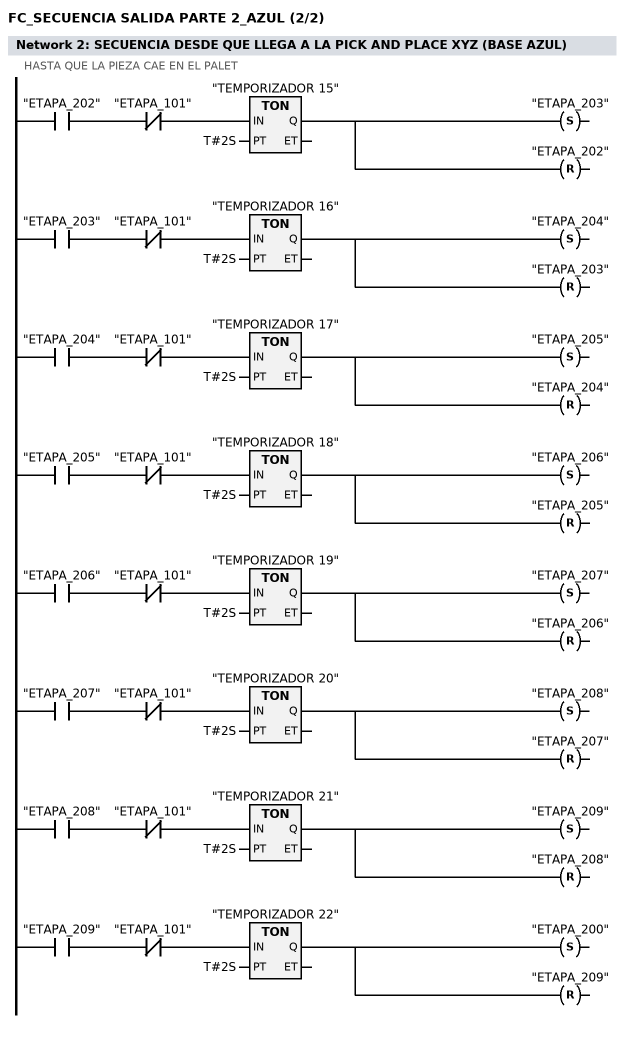
   "TEMPORIZADOR 15".TON(IN := "ETAPA_202" AND NOT "ETAPA_101", PT := T#2S);
   IF "TEMPORIZADOR 15".Q THEN
       "ETAPA_203" := TRUE;
       "ETAPA_202" := FALSE;
   END_IF;
   "TEMPORIZADOR 16".TON(IN := "ETAPA_203" AND NOT "ETAPA_101", PT := T#2S);
   IF "TEMPORIZADOR 16".Q THEN
       "ETAPA_204" := TRUE;
       "ETAPA_203" := FALSE;
   END_IF;
   "TEMPORIZADOR 17".TON(IN := "ETAPA_204" AND NOT "ETAPA_101", PT := T#2S);
   IF "TEMPORIZADOR 17".Q THEN
       "ETAPA_205" := TRUE;
       "ETAPA_204" := FALSE;
   END_IF;
   "TEMPORIZADOR 18".TON(IN := "ETAPA_205" AND NOT "ETAPA_101", PT := T#2S);
   IF "TEMPORIZADOR 18".Q THEN
       "ETAPA_206" := TRUE;
       "ETAPA_205" := FALSE;
   END_IF;
   "TEMPORIZADOR 19".TON(IN := "ETAPA_206" AND NOT "ETAPA_101", PT := T#2S);
   IF "TEMPORIZADOR 19".Q THEN
       "ETAPA_207" := TRUE;
       "ETAPA_206" := FALSE;
   END_IF;
   "TEMPORIZADOR 20".TON(IN := "ETAPA_207" AND NOT "ETAPA_101", PT := T#2S);
   IF "TEMPORIZADOR 20".Q THEN
       "ETAPA_208" := TRUE;
       "ETAPA_207" := FALSE;
   END_IF;
   "TEMPORIZADOR 21".TON(IN := "ETAPA_208" AND NOT "ETAPA_101", PT := T#2S);
   IF "TEMPORIZADOR 21".Q THEN
       "ETAPA_209" := TRUE;
       "ETAPA_208" := FALSE;
   END_IF;
   "TEMPORIZADOR 22".TON(IN := "ETAPA_209" AND NOT "ETAPA_101", PT := T#2S);
   IF "TEMPORIZADOR 22".Q THEN
       "ETAPA_200" := TRUE;
       "ETAPA_209" := FALSE;
   END_IF;
END_REGION
END_FUNCTION

FUNCTION "FC_BOBINAS SALIDA PARTE 2_AZUL" : Void   // FC9, LAD
{ S7_Optimized_Access := 'TRUE' }
VERSION : 0.1
// EN ESTE BLOQUE SE ENCUENTRA LA ASIGNACIÓN DE CADA ETAPA CON EL ACTUADOR QUE CORRESPONDE, DESDE QUE LAS PIEZAS AZULES PASAN LAS CÁMARAS DE VISIÓN DE COLORES HASTA QUE LA PICK&PLACE XYZ LAS DEJA EN EL PALET
BEGIN

REGION Network 1: ASIGNACION BOBINAS A PARTIR DE QUE LAS CÁMARAS DISCRIMINAN(CAMINO BASE AZUL)
   // HASTA QUE LA PICK AND PLACE XYZ DEJA LA BASE AZUL EN EL PALET
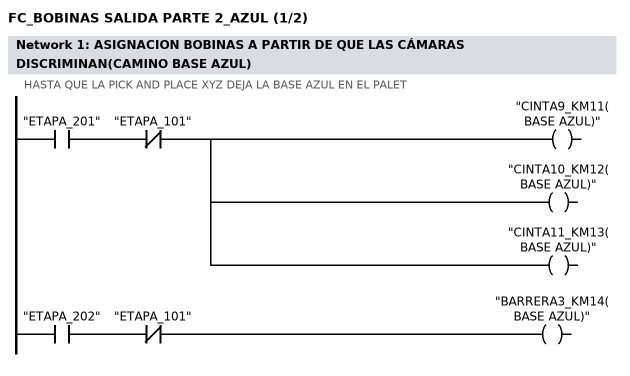
   RUNG wire#powerrail
      Contact( "ETAPA_201" )
      I_Contact( "ETAPA_101" )
      wire#w1
      Coil( "CINTA9_KM11(BASE AZUL)" )
   END_RUNG
   RUNG wire#w1
      Coil( "CINTA10_KM12(BASE AZUL)" )
   END_RUNG
   RUNG wire#w1
      Coil( "CINTA11_KM13(BASE AZUL)" )
   END_RUNG
   RUNG wire#powerrail
      Contact( "ETAPA_202" )
      I_Contact( "ETAPA_101" )
      Coil( "BARRERA3_KM14(BASE AZUL)" )
   END_RUNG
   // the same network as SCL:
   "CINTA9_KM11(BASE AZUL)" := "ETAPA_201" AND NOT "ETAPA_101";
   "CINTA10_KM12(BASE AZUL)" := "CINTA9_KM11(BASE AZUL)";
   "CINTA11_KM13(BASE AZUL)" := "CINTA9_KM11(BASE AZUL)";
   "BARRERA3_KM14(BASE AZUL)" := "ETAPA_202" AND NOT "ETAPA_101";
END_REGION

REGION Network 2: ASIGNACION BOBINAS DESDE QUE LLEGA A LA PICK AND PLACE XYZ (BASE AZUL)
   // HASTA QUE LA PIEZA CAE EN EL PALET
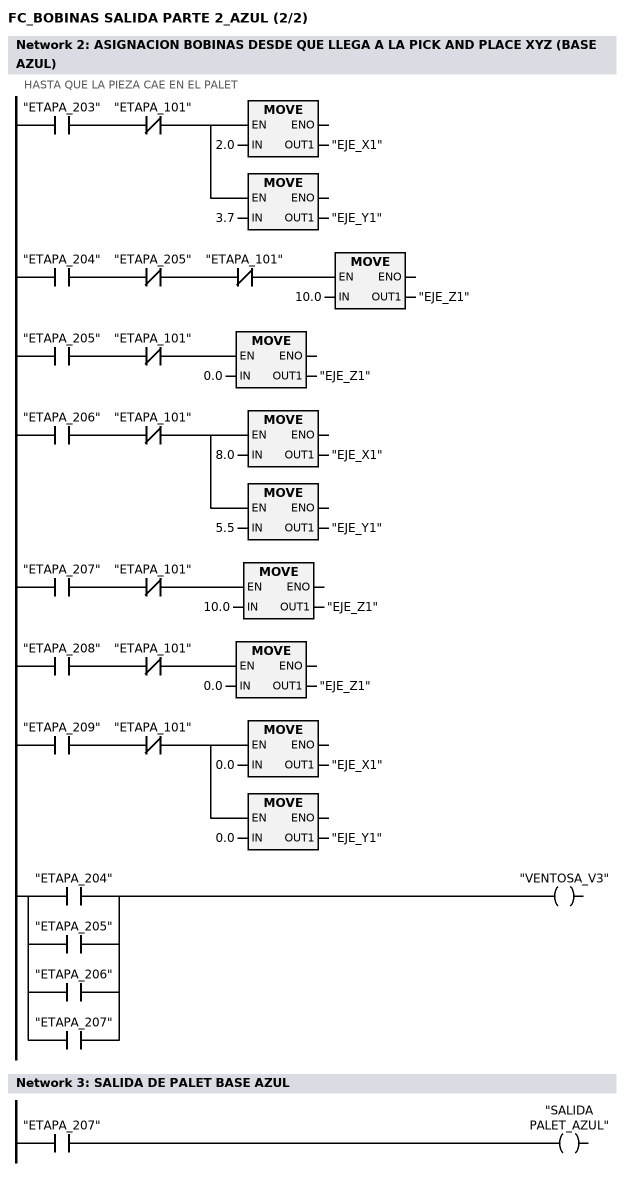
   RUNG wire#powerrail
      Contact( "ETAPA_203" )
      I_Contact( "ETAPA_101" )
      wire#w1
      Move(in := 2.0, out1 => "EJE_X1")
   END_RUNG
   RUNG wire#w1
      Move(in := 3.7, out1 => "EJE_Y1")
   END_RUNG
   RUNG wire#powerrail
      Contact( "ETAPA_204" )
      I_Contact( "ETAPA_205" )
      I_Contact( "ETAPA_101" )
      Move(in := 10.0, out1 => "EJE_Z1")
   END_RUNG
   RUNG wire#powerrail
      Contact( "ETAPA_205" )
      I_Contact( "ETAPA_101" )
      Move(in := 0.0, out1 => "EJE_Z1")
   END_RUNG
   RUNG wire#powerrail
      Contact( "ETAPA_206" )
      I_Contact( "ETAPA_101" )
      wire#w2
      Move(in := 8.0, out1 => "EJE_X1")
   END_RUNG
   RUNG wire#w2
      Move(in := 5.5, out1 => "EJE_Y1")
   END_RUNG
   RUNG wire#powerrail
      Contact( "ETAPA_207" )
      I_Contact( "ETAPA_101" )
      Move(in := 10.0, out1 => "EJE_Z1")
   END_RUNG
   RUNG wire#powerrail
      Contact( "ETAPA_208" )
      I_Contact( "ETAPA_101" )
      Move(in := 0.0, out1 => "EJE_Z1")
   END_RUNG
   RUNG wire#powerrail
      Contact( "ETAPA_209" )
      I_Contact( "ETAPA_101" )
      wire#w3
      Move(in := 0.0, out1 => "EJE_X1")
   END_RUNG
   RUNG wire#w3
      Move(in := 0.0, out1 => "EJE_Y1")
   END_RUNG
   RUNG wire#powerrail
      Contact( "ETAPA_204" )
      wire#w4
      Coil( "VENTOSA_V3" )
   END_RUNG
   RUNG wire#powerrail
      Contact( "ETAPA_205" )
   END_RUNG wire#w4
   RUNG wire#powerrail
      Contact( "ETAPA_206" )
   END_RUNG wire#w4
   RUNG wire#powerrail
      Contact( "ETAPA_207" )
   END_RUNG wire#w4
   // the same network as SCL:
   IF "ETAPA_203" AND NOT "ETAPA_101" THEN
       "EJE_X1" := 2.0;
       "EJE_Y1" := 3.7;
   END_IF;
   IF "ETAPA_204" AND NOT "ETAPA_205" AND NOT "ETAPA_101" THEN "EJE_Z1" := 10.0; END_IF;
   IF "ETAPA_205" AND NOT "ETAPA_101" THEN "EJE_Z1" := 0.0; END_IF;
   IF "ETAPA_206" AND NOT "ETAPA_101" THEN
       "EJE_X1" := 8.0;
       "EJE_Y1" := 5.5;
   END_IF;
   IF "ETAPA_207" AND NOT "ETAPA_101" THEN "EJE_Z1" := 10.0; END_IF;
   IF "ETAPA_208" AND NOT "ETAPA_101" THEN "EJE_Z1" := 0.0; END_IF;
   IF "ETAPA_209" AND NOT "ETAPA_101" THEN
       "EJE_X1" := 0.0;
       "EJE_Y1" := 0.0;
   END_IF;
   "VENTOSA_V3" := "ETAPA_204" OR "ETAPA_205" OR "ETAPA_206" OR "ETAPA_207";
END_REGION

REGION Network 3: SALIDA DE PALET BASE AZUL
   RUNG wire#powerrail
      Contact( "ETAPA_207" )
      Coil( "SALIDA PALET_AZUL" )
   END_RUNG
   // the same network as SCL:
   "SALIDA PALET_AZUL" := "ETAPA_207";
END_REGION
END_FUNCTION

FUNCTION "FC_SECUENCIA SALIDA PARTE 2_VERDE" : Void   // FC10, LAD
{ S7_Optimized_Access := 'TRUE' }
VERSION : 0.1
// EN ESTE BLOQUE SE ENCUENTRA LA PROGRAMACIÓN DE LA SECUENCIA DESDE QUE LAS CÁMARAS DE VISION DE COLORES DISCRIMAN LA PIEZA VERDE HASTA QUE LA PICK&PLACE XYZ LAS DEJA EN UN PALET
BEGIN

REGION Network 1: SECUENCIA DEL PROCESO DE SALIDA PARTE 2(CAMINO BASE VERDE)
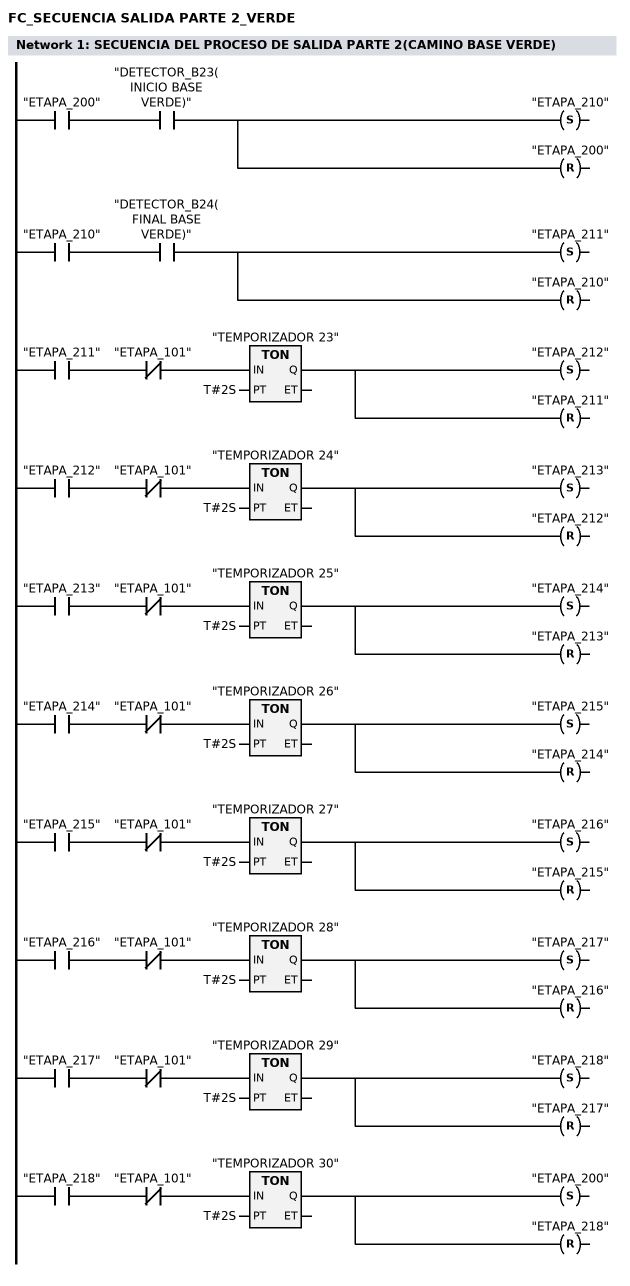
   IF "ETAPA_200" AND "DETECTOR_B23(INICIO BASE VERDE)" THEN
       "ETAPA_210" := TRUE;
       "ETAPA_200" := FALSE;
   END_IF;
   IF "ETAPA_210" AND "DETECTOR_B24(FINAL BASE VERDE)" THEN
       "ETAPA_211" := TRUE;
       "ETAPA_210" := FALSE;
   END_IF;
   "TEMPORIZADOR 23".TON(IN := "ETAPA_211" AND NOT "ETAPA_101", PT := T#2S);
   IF "TEMPORIZADOR 23".Q THEN
       "ETAPA_212" := TRUE;
       "ETAPA_211" := FALSE;
   END_IF;
   "TEMPORIZADOR 24".TON(IN := "ETAPA_212" AND NOT "ETAPA_101", PT := T#2S);
   IF "TEMPORIZADOR 24".Q THEN
       "ETAPA_213" := TRUE;
       "ETAPA_212" := FALSE;
   END_IF;
   "TEMPORIZADOR 25".TON(IN := "ETAPA_213" AND NOT "ETAPA_101", PT := T#2S);
   IF "TEMPORIZADOR 25".Q THEN
       "ETAPA_214" := TRUE;
       "ETAPA_213" := FALSE;
   END_IF;
   "TEMPORIZADOR 26".TON(IN := "ETAPA_214" AND NOT "ETAPA_101", PT := T#2S);
   IF "TEMPORIZADOR 26".Q THEN
       "ETAPA_215" := TRUE;
       "ETAPA_214" := FALSE;
   END_IF;
   "TEMPORIZADOR 27".TON(IN := "ETAPA_215" AND NOT "ETAPA_101", PT := T#2S);
   IF "TEMPORIZADOR 27".Q THEN
       "ETAPA_216" := TRUE;
       "ETAPA_215" := FALSE;
   END_IF;
   "TEMPORIZADOR 28".TON(IN := "ETAPA_216" AND NOT "ETAPA_101", PT := T#2S);
   IF "TEMPORIZADOR 28".Q THEN
       "ETAPA_217" := TRUE;
       "ETAPA_216" := FALSE;
   END_IF;
   "TEMPORIZADOR 29".TON(IN := "ETAPA_217" AND NOT "ETAPA_101", PT := T#2S);
   IF "TEMPORIZADOR 29".Q THEN
       "ETAPA_218" := TRUE;
       "ETAPA_217" := FALSE;
   END_IF;
   "TEMPORIZADOR 30".TON(IN := "ETAPA_218" AND NOT "ETAPA_101", PT := T#2S);
   IF "TEMPORIZADOR 30".Q THEN
       "ETAPA_200" := TRUE;
       "ETAPA_218" := FALSE;
   END_IF;
END_REGION
END_FUNCTION

FUNCTION "FC_BOBINAS SALIDA PARTE 2_VERDE" : Void   // FC11, LAD
{ S7_Optimized_Access := 'TRUE' }
VERSION : 0.1
// EN ESTE BLOQUE SE ENCUENTRA LA ASIGNACIÓN DE CADA ETAPA CON EL ACTUADOR QUE CORRESPONDE, DESDE QUE LAS PIEZAS VERDES PASAN LAS CÁMARAS DE VISIÓN DE COLORES HASTA QUE LA PICK&PLACE XYZ LAS DEJA EN EL PALET
BEGIN

REGION Network 1: ASIGNACION BOBINAS A PARTIR DE QUE LAS CÁMARAS DISCRIMINAN(CAMINO BASE VERDE)
